(* IEC 61131-3 sources: daoli-st-library/DL_Process (part 40) *)

(* ---- FB_DL_LineChangeoverChecklist.st ---- *)
(*==============================================================================
 * 组件名称 (Component)  : FB_DL_LineChangeoverChecklist
 * 溯源说明 (Provenance) : 道莅 clean-room 防御性实现（PackML 深化）
 * 所属子库 (Sublibrary) : DL_Process / Changeover
 * 当前版本 (Version)    : 1.0.1
 * 兼容性   (Platform)   : CODESYS 3.5 / TwinCAT 3 / 汇川 InoProShop；
 *                         纯 IEC 61131-3（第 3 版），零标准库依赖
 * 组件分类 (Category)   : 功能块（FUNCTION_BLOCK）· 换型检查清单顺控
 * 功能一句话 (Summary)  : 检查项逐步确认 + 前向跳步登记 + 未完成禁止启动。
 * 边界与安全 (Boundary) : ①跳步仅允许前向（不小于当前步）且不可跳最后一项；
 *                         ②未全部完成（含已跳步）时启动确认拒绝并置码 0362；
 *                         ③回退方向跳步申请拒绝并置码 0361；
 *                         ④bReset 清跳步登记与状态（已完成位由调用方维护）；
 *                         ⑤数组下标全程钳位（禁越界访问）。
 * 错误码    : 16#0005_0361 非法回退跳步申请——信息级（单拍）
 *             16#0005_0362 未完成启动尝试（启动确认被拒）——故障级（单拍）
 * 码位总账  : 16#0005_0361 用 / 16#0005_0362 用
 * 修改记录  : v1.0.0 R26 初版
 *             v1.0.1 R26 终审修复：跳步登记循环补双表异界防御——abSkipReq 与
 *             abStepsDone 为两张独立 ARRAY[*]，申请表更长时按自身 UPPER_BOUND 判界
 *==============================================================================*)
TYPE E_DL_ChgoverState :
(
    eIdle     := 0, // 空闲：未开始检查 / Idle: checklist not started
    eRunning  := 1, // 检查中：存在未确认项 / Running: items pending
    eAllDone  := 2  // 全部完成：允许启动 / All done: start permitted
);
END_TYPE

FUNCTION_BLOCK FB_DL_LineChangeoverChecklist
VAR_INPUT
    abSkipReq     : ARRAY[*] OF BOOL; // 跳步申请位表（与完成位同界）/ Skip request bits
    bStartConfirm : BOOL; // 启动确认请求 / Start confirmation request
    bReset        : BOOL; // 复位：清跳步与状态 / Reset: clear skips and state
END_VAR
VAR_IN_OUT
    abStepsDone : ARRAY[*] OF BOOL; // 检查项完成位表 / Checklist done bits
END_VAR
VAR_OUTPUT
    eState    : E_DL_ChgoverState; // 清单状态机状态 / Checklist state machine state
    uCurStep  : UINT;  // 当前待确认步序号 / Current pending step index
    bAllDone  : BOOL;  // 全部完成（含跳步）/ All done including skips
    bSkipUsed : BOOL;  // 本轮发生过跳步 / Any skip used this round
    eErr      : UDINT; // 本周期错误码，0=无错 / Error code this cycle, 0 = none
END_VAR
VAR
    nSteps  : INT;  // 总步数 / Total step count
    i       : INT;  // 扫描游标 / Scan cursor
    iCur    : INT;  // 当前待确认步内部值 / Current pending step internal
    bPending: BOOL; // 存在未确认项 / Any item pending
    rSkip   : R_TRIG; // 跳步申请沿检测（无条件刷新）/ Skip request edge
    bAnyReq : BOOL; // 跳步申请或哨兵 / Skip request or sentinel
    bUndone : BOOL; // 完成位安全读取副本（双表异界防御）/ Safe done-bit read copy
END_VAR

// ---------- 无条件周期刷新：跳步沿检测（哨兵时钟法，单实例单调用） ----------
bAnyReq := FALSE;
FOR i := 0 TO UPPER_BOUND(abSkipReq, 1) DO
    IF abSkipReq[i] THEN
        bAnyReq := TRUE;                      // 任一跳步申请 / Any skip requested
    END_IF
END_FOR
rSkip(CLK := bAnyReq);

// ---------- 复位：清跳步登记与状态 ----------
IF bReset THEN
    bSkipUsed := FALSE;                       // 跳步登记清零 / Skip ledger cleared
    eState := E_DL_ChgoverState.eIdle;        // 回空闲 / Back to idle
    eErr := 0;
END_IF

// ---------- 周期起点：错误码先清（单拍码生命周期） ----------
eErr := 0;

// ---------- 步数与界防御 ----------
nSteps := UPPER_BOUND(abStepsDone, 1) + 1;    // 总步数 / Total steps
IF nSteps < 1 THEN
    nSteps := 1;                              // 下限防御 / Lower bound guard
END_IF

// ---------- 跳步登记：仅前向且不可跳最后一项 ----------
IF rSkip.Q THEN
    FOR i := 0 TO UPPER_BOUND(abSkipReq, 1) DO
        // 双表异界防御：完成位读取按 abStepsDone 自身上界判界 / Bounds guard for mismatched tables
        IF i <= UPPER_BOUND(abStepsDone, 1) THEN
            bUndone := NOT abStepsDone[i];    // 完成位安全读取 / Safe done-bit read
        ELSE
            bUndone := FALSE;                 // 越界位视作不可登记 / Out-of-range: not registrable
        END_IF
        IF abSkipReq[i] AND bUndone AND (i < nSteps - 1) THEN
            // 前向且非最后一项：跳步视同完成登记（台账语义）/ Forward & not last: mark done
            abStepsDone[i] := TRUE;           // 跳步登记 / Skip marks done
            bSkipUsed := TRUE;                // 记录跳步 / Skip recorded
        ELSIF abSkipReq[i] AND bUndone AND (i >= nSteps - 1) THEN
            eErr := 16#0005_0361;             // 末项禁跳码 / Last-step skip forbidden
        END_IF
    END_FOR
END_IF

// ---------- 当前步扫描：首个未确认项（下标钳位） ----------
iCur := 0;
bPending := FALSE;
FOR i := 0 TO nSteps - 1 DO
    IF NOT abStepsDone[i] THEN
        iCur := i;                            // 首个未确认项 / First pending item
        bPending := TRUE;                     // 存在未确认 / Pending exists
        EXIT;                                 // 找到即出（最小编号优先）/ Exit on first
    END_IF
END_FOR
uCurStep := INT_TO_UINT(iCur);                // 对外当前步 / Exposed current step

// ---------- 状态机：CASE 覆盖全部枚举成员加 ELSE 兜底 ----------
CASE eState OF
    E_DL_ChgoverState.eIdle:                  // 拍 N 进入：空闲 / Entered: idle
        IF bPending THEN
            eState := E_DL_ChgoverState.eRunning; // 有未确认项进检查态 / Pending found, running
        END_IF
        // 本拍行为：空闲等待 / This cycle: idle waiting
        // 拍 N+1 转出：进 eRunning / Leaving to running

    E_DL_ChgoverState.eRunning:               // 拍 N 进入：检查中 / Entered: running
        IF NOT bPending THEN
            eState := E_DL_ChgoverState.eAllDone; // 全确认进完成态 / All confirmed, done
        END_IF
        // 本拍行为：保持当前步等待确认 / This cycle: hold current step
        // 拍 N+1 转出：eAllDone 或保持 / Leaving to done or hold

    E_DL_ChgoverState.eAllDone:               // 拍 N 进入：全部完成 / Entered: all done
        bAllDone := TRUE;                     // 放行启动 / Permit start
        IF bPending THEN
            eState := E_DL_ChgoverState.eRunning; // 调用方清位后回检查态 / Back to running
        END_IF
        // 本拍行为：保持放行 / This cycle: keep permit
        // 拍 N+1 转出：条件驱动 / Condition-driven leaving

    ELSE                                      // 非法状态兜底回空闲 / Illegal state fallback
        eState := E_DL_ChgoverState.eIdle;
        bAllDone := FALSE;
END_CASE

// ---------- bAllDone 与状态同步（保持单口径） ----------
IF eState = E_DL_ChgoverState.eAllDone THEN
    bAllDone := TRUE;
ELSE
    bAllDone := FALSE;                        // 非完成态不放行 / No permit unless done
END_IF

// ---------- 启动确认仲裁：未全部完成拒绝 ----------
IF bStartConfirm AND (NOT bAllDone) THEN
    eErr := 16#0005_0362;                     // 未完成启动尝试码 / Start attempt while incomplete
END_IF

END_FUNCTION_BLOCK

(* ---- FB_DL_LineClearanceVerify.st ---- *)
(*
  ==================================================================
  组件名 Component  : FB_DL_LineClearanceVerify
  分类   Category   : DL_Process
  前缀   Naming     : FB_DL_ ｜ b/n/u/f/t/e/st 类型前缀制（R265）
  复杂度 Complexity  : 高
  版本   Version    : 1.0.1
  功能   Purpose    : 换型清线验证（清料确认 + 残留计数 + 阶段确认窗状态机 + 超窗升级码）。
  来源   Source     : self-std（换型清线公开工艺语义自研）
  平台   Platform   : 纯 IEC 61131-3（TON / R_TRIG / CASE），三平台通用
  分工声明 Split     : 与 FB_DL_ChangeoverSequence（换型顺控属主）与
                      FB_DL_ShiftHandoverCheck（交接检查属主）分工——本件只做
                      换型时点的清线验证闭环（R216 双向互引）。
  作者   Author     : 道莅代码库 · PLC 编程专家（R61）
  归属 Ownership     : E_DL_ClearPhase 属主为本文件（全库唯一定义，R264）；
                      引用件只引用不重声明。
  ------------------------------------------------------------------
  边界 Boundary     :
                      一 残留计数清零判据用整数精确比较（uResidueCnt = 0，禁浮点）；
                      二 同拍竞态先消化确认沿再判超窗（R275 模板：段 3 预消化
                         确认沿，段 4 才判窗口到期迁移）；
                      三 快照/计数出口纳入复位清单（R243）：复位沿清残留计数、
                         清阶段计数与迁相位（R311 作用域逐项声明）；
                      四 组态窗非法（tConfirmWin ≤ 0 或 nResidueMax < 0）判故障
                         锁存（3038）；超窗升级独立码 3037（R190 归因唯一）；
                      五 CASE 必带 ELSE 兜底；TON/R_TRIG 段 0 无条件刷新（R7），
                         TON IN 串故障锁存门控（FB50-1）；
                      六 无全局、无外部变量、无物理地址。
  错误码   Codes    :
    16#0005_3036【信息级】清线确认窗内残留计数超过 nResidueMax 时逐拍提示
                            （默认 0 = 残留非零即提示）；不锁存、不置 bError、
                            不阻断放行（口径以实现为准，v1.0.1 注释订正）
    16#0005_3037【故障级】阶段确认窗到期仍未确认，升级锁存至复位沿
    16#0005_3038【故障级】组态非法（确认窗 ≤ 0 或残留上限 < 0），锁存至复位沿
  码位口径   Code Note :
    3036 为信息级，在段 5 的 ELSIF 链中固定排于故障回放之后（链末位），
    故故障相下 3036 不可能覆盖已置的故障码（R190 归因唯一 + R285 分级纪律）；
    3036 逐拍重算不锁存，残留计数回落至上限以内即自动消失。
  验收   Acceptance :
    算法已证（脚本）：未跑 ｜ 编译器已证（三平台）：未跑
    V1 无残留、窗内确认沿 → bClearOk 单拍、无故障
    V2 残留 3 件逐件出清后确认 → 计数 3、bClearOk 单拍
    V3 窗到期未确认 → 码 3037、eFault、锁存待复位
    V4 nResidueMax=0、残留 1 件 → eErr=3036、bError=FALSE（信息级不置故障）
    V5 nResidueMax=3、残留 2 件 → eErr=0（允许残留）；残留 4 件 → 3036
    V6 窗非法（tConfirmWin ≤ 0）且残留超限 → 3038 优先，3036 不覆盖
  修订记录 Revision  :
    2026-11-21  v1.0.0  R61 首版（批 4 · 序号 16）
    2026-11-21  v1.0.1  R62-D6 返修：①头注释 3036 口径订正为「确认窗内残留超 nResidueMax 逐拍提示（默认 0 = 非零即提示）；不锁存、不置 bError、不阻断放行」；②引脚注释补默认语义；③复核 3036 在 ELSIF 链末位不覆盖故障码（行为零变更）
  ==================================================================
*)
TYPE E_DL_ClearPhase :
(
    eIdle     := 0,  // 空闲：等清线请求沿 / idle, waiting for the clearance request edge
    eSweep    := 10, // 清料相：残留逐件出清 / the sweeping phase, the residues leaving one by one
    eConfirm  := 20, // 确认相：阶段确认窗内等确认沿 / the confirm phase inside the window
    eFault    := 30  // 故障：超窗或组态非法，锁存待复位 / fault, the overrun or the illegal configuration latched
);
END_TYPE

FUNCTION_BLOCK FB_DL_LineClearanceVerify
VAR_INPUT
    bClearReq    : BOOL := FALSE;  // 清线请求电平，上升沿发起 / the clearance request level
    bItemOut     : BOOL := FALSE;  // 出料口有料电平 [-] / the item present level at the outlet
    bClearConfirm: BOOL := FALSE;  // 清线确认电平，上升沿确认 / the clearance confirm level
    bReset       : BOOL := FALSE;  // 故障复位电平，上升沿清锁存 / the fault reset level
    tConfirmWin  : TIME := T#60S;  // 阶段确认窗时长 [毫秒] / the confirm window duration
    nResidueMax  : DINT := 0;      // 残留计数上限 [件]，≥ 0；默认 0 即残留非零即提示，调大则该量残留仍允许放行 / the residue count bound, non negative; zero means any residue hints, a larger bound tolerates that many residues
END_VAR
VAR_OUTPUT
    uResidueCnt : UDINT := 0;              // 本轮残留计数 [件] / the residue count of this round
    bClearOk    : BOOL := FALSE;           // 清线通过单拍脉冲 [-] / the clearance passed one shot pulse
    eState      : E_DL_ClearPhase;         // 主状态机当前态 [状态] / the current state
    bError      : BOOL := FALSE;           // 故障锁存位（与锁存同源，R191）/ the fault bit from the latch
    eErr        : UDINT := 16#0000_0000;   // 错误码，0 = 正常 / the error code, zero is ok
END_VAR
VAR
    _bInit     : BOOL := FALSE;                            // 首拍初始化标志（R310）/ the first scan flag
    _eState    : E_DL_ClearPhase := E_DL_ClearPhase.eIdle; // 内部状态寄存器 / the internal state register
    _bFault    : BOOL := FALSE;                            // 故障锁存副本（仅复位沿清除）/ the fault latch copy
    _bCfgBad   : BOOL := FALSE;                            // 组态非法标记（逐拍重算入锁存）/ the configuration fault flag
    _uResidue  : UDINT := 0;                               // 残留计数副本 [件] / the residue count copy
    _bOk       : BOOL := FALSE;                            // 通过单拍内部位，段 1 预清段 5 映射 / the internal ok bit
    _bEvtTaken : BOOL := FALSE;                            // 本拍确认沿已消化标记（R275）/ the confirm edge consumed flag
    _bCfgLatch : BOOL := FALSE;                            // 组态锁存副本（与 _bCfgBad 区分：锁存型）/ the configuration latch copy
    rtReq      : R_TRIG;  // 清线请求沿实例，段 0 无条件刷新 / the request edge instance
    rtItem     : R_TRIG;  // 出料沿实例，段 0 无条件刷新 / the item out edge instance
    rtConfirm  : R_TRIG;  // 确认沿实例，段 0 无条件刷新 / the confirm edge instance
    rtReset    : R_TRIG;  // 复位沿实例，段 0 无条件刷新 / the reset edge instance
    tonWin     : TON;     // 阶段确认窗定时器，段 0 无条件刷新 / the confirm window timer
END_VAR

// 段 0｜定时器与沿检测无条件周期刷新（禁入分支，R7；TON IN 串故障锁存门控，FB50-1）/ segment 0, the unconditional refresh
rtReq(CLK := bClearReq); // 请求沿 / the request edge
rtItem(CLK := bItemOut); // 出料沿 / the item out edge
rtConfirm(CLK := bClearConfirm); // 确认沿 / the confirm edge
rtReset(CLK := bReset); // 复位沿 / the reset edge
tonWin(IN := (_eState = E_DL_ClearPhase.eConfirm) AND (NOT _bFault), PT := tConfirmWin); // 确认窗：仅确认相且无锁存时计时 / the window timing only in the confirm phase

// 段 1｜首拍初始化与单拍标志预清（R310 / FB32-1 / R256）/ segment 1, the first scan init and the preset
IF NOT _bInit THEN // 首拍一拍 / the first scan
    _bInit := TRUE; // 置首拍标志 / raise the first scan flag
    _bFault := FALSE; // 故障锁存显式清零 / clear the fault latch explicitly
    _bCfgLatch := FALSE; // 组态锁存显式清零 / clear the configuration latch explicitly
    _uResidue := 0; // 残留计数显式清零 / clear the residue count explicitly
    _eState := E_DL_ClearPhase.eIdle; // 状态显式落空闲 / place the state to idle
END_IF
IF rtReset.Q THEN // 复位沿（作用域：清锁存 + 清计数 + 迁相位，R311 / R243 声明）/ the reset edge with the declared scope
    _bFault := FALSE; // 清故障锁存（解除路径：复位沿恒可达，R152 自证）/ clear the fault latch
    _bCfgLatch := FALSE; // 清组态锁存 / clear the configuration latch
    _uResidue := 0; // 清残留计数（R243 快照/计数出口入复位清单）/ clear the residue count
    _eState := E_DL_ClearPhase.eIdle; // 迁回空闲 / back to idle
END_IF
_bOk := FALSE; // 通过单拍预清零 / preset the ok bit false
_bEvtTaken := FALSE; // 确认沿消化标记预清零 / preset the consumed flag false
_bCfgBad := FALSE; // 组态标记预清零 / preset the configuration flag false

// 段 2｜组态域闸（边界四）/ segment 2, the configuration gate
IF (tConfirmWin <= T#0S) OR (nResidueMax < 0) THEN // 窗非法或上限负 / an illegal window or a negative bound
    _bCfgBad := TRUE; // 置组态标记 / raise the configuration flag
    _bCfgLatch := TRUE; // 锁存组态故障（3038）/ latch the configuration fault
    _bFault := TRUE; // 总锁存（段 4 迁移）/ latch the total fault
END_IF

// 段 3｜本拍确认沿预消化（R275：合法事件先于窗口到期迁移消化）/ segment 3, the confirm edge pre digest
IF rtConfirm.Q AND (_eState = E_DL_ClearPhase.eConfirm) AND (NOT _bFault) THEN // 确认相内的确认沿 / a confirm edge inside the confirm phase
    _bEvtTaken := TRUE; // 标记本拍已消化（段 4 不再判超窗）/ mark the edge consumed this scan
    _bOk := TRUE; // 置通过单拍 / raise the ok bit
    _eState := E_DL_ClearPhase.eIdle; // 迁回空闲（本轮通过）/ back to idle with the round passed
END_IF

// 段 4｜主状态机（ENUM + CASE，ELSE 兜底；超窗迁移让位于本拍确认沿，边界二）/ segment 4, the main machine
CASE _eState OF
    E_DL_ClearPhase.eIdle: // 空闲相 / the idle phase
        IF rtReq.Q AND (NOT _bFault) THEN // 请求沿 + 闸位复检（R274）/ the request edge with the gate recheck
            _uResidue := 0; // 新一轮残留计数归零（整数精确） / reset the residue count by the exact integer
            _eState := E_DL_ClearPhase.eSweep; // 迁入清料相 / enter the sweeping phase
        END_IF
    E_DL_ClearPhase.eSweep: // 清料相：残留逐件出清 / the sweeping phase
        IF rtItem.Q THEN // 出料沿：残留计一件 / an item out edge counts one residue
            _uResidue := _uResidue + 1; // 残留计数推进 / advance the residue count
        END_IF
        IF (NOT bItemOut) AND (NOT rtItem.Q) THEN // 出料口已空且本拍无新出料沿（整数域判据，边界一）/ the outlet empty with no new edge
            _eState := E_DL_ClearPhase.eConfirm; // 迁入确认相（确认窗起算）/ enter the confirm phase
        ELSIF _bFault THEN // 前置条件消失出口 / the prerequisite gone exit
            _eState := E_DL_ClearPhase.eFault; // 迁入故障相 / enter the fault phase
        END_IF
    E_DL_ClearPhase.eConfirm: // 确认相（本拍确认沿已在段 3 消化并迁出，边界二）/ the confirm phase, the edge already digested in segment three
        IF tonWin.Q AND (NOT _bEvtTaken) THEN // 窗口到期且本拍无确认沿（R275 同拍竞态口径）/ the window expired with no confirm edge this scan
            _bFault := TRUE; // 锁存超窗故障（3037，升级码）/ latch the overrun fault
        ELSIF _bFault THEN // 前置条件消失 / the prerequisite gone
            _eState := E_DL_ClearPhase.eFault; // 迁入故障相 / enter the fault phase
        END_IF
    E_DL_ClearPhase.eFault: // 故障相：等复位沿（解除可达，边界三）/ the fault phase until the reset
        IF NOT _bFault THEN // 锁存已清才迁出（防清锁同拍重锁，FB50-1）/ the exit after the latch cleared
            _eState := E_DL_ClearPhase.eIdle; // 迁回空闲 / back to idle
        END_IF
    ELSE // 非法枚举值拦截 / the illegal enumeration guard
        _eState := E_DL_ClearPhase.eIdle; // 落回空闲 / force back to idle
        _bFault := TRUE; // 置锁存 / latch the fault
END_CASE

// 段 5｜统一出口（内部副本单点映射；故障码锁存回放，R187）/ segment 5, the unified outlet
uResidueCnt := _uResidue; // 残留计数出口 / the residue count outlet
bClearOk := _bOk; // 通过单拍出口 / the ok pulse outlet
eState := _eState; // 状态出口 / the state outlet
bError := _bFault; // 故障位出口（与锁存同源）/ the fault bit outlet
IF _bFault THEN // 故障锁存回放优先 / the latched fault replays first
    IF _bCfgLatch THEN // 组态成因（独立码值，R190）/ the configuration cause
        eErr := 16#0005_3038; // 故障级：组态非法 / fault grade, the illegal configuration
    ELSE // 超窗成因 / the overrun cause
        eErr := 16#0005_3037; // 故障级：确认窗到期未确认，升级 / fault grade, the overrun escalated
    END_IF
ELSIF (_uResidue > DINT_TO_UDINT(nResidueMax)) OR (nResidueMax < 0) THEN // 残留超限提示（信息级，排在故障回放之后即链末位，不覆盖故障码，R285）/ the residue over the bound, informational and last in the chain so it never covers a fault code
    eErr := 16#0005_3036; // 信息级：残留计数非零超提示限 / informational, the residues over the hint bound
ELSE // 无事件 / no event
    eErr := 16#0000_0000; // 正常 / ok
END_IF
END_FUNCTION_BLOCK

(* ---- FB_DL_LoadlockPressureCross.st ---- *)
(*
  FB_DL_LoadlockPressureCross  —  Loadlock 双表压力交叉校验与误开门拦截 / Loadlock dual-gauge cross check and door interlock
  分类 Category : DL_Process
  码位 Code     : 16#06_0_83
  版本 Version  : 1.0.0
  溯源 Source   : ISA-18.2 语义借鉴 · clean-room 实现，仅借分类/参数域/命名，未复制源码
  功能 Function : 1) 双表压力各自过 NE43 有效域后计算偏差，偏差越窗即判交叉故障并锁存首出表号；
                  2) 任一表无效即禁开门（禁用无效值参与偏差计算）；
                  3) 开门许可仅由「双表一致 AND 压力到位」两条件同时满足产生，解除路径可达。
  边界 Boundary : ① 双表各自 NE43 有效域闸，任一无效即禁开门，禁用无效值参与偏差计算；
                  ② 偏差窗上下限配比约束（容差 > 0、目标压力 > 0、迟滞 ≤ 容差/2），非法即组态报码；
                  ③ 许可解锁条件可从「双表一致 AND 压力到位」到达（FB33-2 可达性）；
                  ④ 拦截态三行同向：许可 FALSE → 偏差记录保持 → 拦截标志 TRUE。
  依赖 Depends  : FB_DL_ToleranceWindow（偏差窗判定，每拍无条件调用）

  码表 Error codes（本件子码步进 16#10，避让邻件码位）:
    16#0002_0683 故障级：偏差窗组态非法（容差 <= 0 或迟滞 > 容差/2 或目标压力 <= 0）
    16#0002_0693 故障级：表 A / 表 B 信号无效（NE43 域外或缺省），禁开门
    16#0002_06A3 信息级：交叉偏差越窗（信息记录，故障锁存由 0683 族承担）
*)

TYPE E_DL_LlxcPhase :
(
    eIdle    := 0,   // 空闲 / Idle
    eCheck   := 10,  // 偏差校验中 / Cross check running
    ePermit  := 20,  // 允许开门 / Door permitted
    eBlocked := 30,  // 拦截（表无效或偏差越窗）/ Blocked
    eFault   := 90   // 故障锁定 / Fault locked
);
END_TYPE

FUNCTION_BLOCK FB_DL_LoadlockPressureCross
VAR_INPUT
    bEnable       : BOOL;                         // 总使能，FALSE 禁开门 / Master enable, FALSE forbids door
    bReset        : BOOL;                         // 复位，上升沿清锁存 / Reset, clears latches
    fPressAKPa    : REAL;                         // 表 A 压力 [kPa abs]，域 0.001~200 / Gauge A pressure [kPa abs]
    bValidAK      : BOOL;                         // 表 A 信号有效（NE43 已在传感器侧判定）/ Gauge A signal valid
    fPressBKPa    : REAL;                         // 表 B 压力 [kPa abs]，域 0.001~200 / Gauge B pressure [kPa abs]
    bValidBK      : BOOL;                         // 表 B 信号有效 / Gauge B signal valid
    fDevMaxKPa    : REAL := 0.5;                  // 允许交叉偏差 [kPa]，域 > 0 / Allowed cross deviation [kPa]
    fDevHystKPa   : REAL := 0.05;                 // 偏差窗迟滞 [kPa]，域 0~容差/2 / Deviation hysteresis [kPa]
    fPressTargetKPa : REAL := 101.3;              // 开门目标压力 [kPa abs]，域 > 0 / Door-open target pressure
    fPressTolKPa  : REAL := 5.0;                  // 压力到位容差 [kPa]，域 > 0 / Pressure-in-place tolerance
    fEps          : REAL := 1.0E-6;               // 浮点判零容差 [1] / Floating zero tolerance
END_VAR
VAR_OUTPUT
    bDoorPermit   : BOOL;                         // 开门许可（唯一放行信号）/ Door permit, the only release
    bCrossFault   : BOOL;                         // 交叉故障标志（保持型）/ Cross fault flag, held
    bPressInPlace : BOOL;                         // 压力到位标志 / Pressure in place
    fDevKPa       : REAL;                         // 当前双表偏差 [kPa] / Current cross deviation [kPa]
    nFirstOut     : INT;                          // 首出表号 1 = A，2 = B，0 = 无 / First-out gauge, 0 = none
    bError        : BOOL;                         // 故障标志，与故障级码配对 / Fault flag paired with fault codes
    uErrorId      : UDINT;                        // 事件码，0 = 无事件 / Event code, 0 = none
    eStateOut     : E_DL_LlxcPhase;               // 状态机当前态，段尾单点映射 / Phase mapped at tail
END_VAR
VAR
    _eState       : E_DL_LlxcPhase := E_DL_LlxcPhase.eIdle;  // 内部状态 / Internal state
    rtrReset      : R_TRIG;                       // 复位沿 / Reset edge
    fbDevWin      : FB_DL_ToleranceWindow;        // 偏差窗判定实例（无条件调用）/ Deviation window instance
    bCfgOk        : BOOL;                         // 组态合法标志 / Configuration valid
    bAOk          : BOOL;                         // 表 A 有效（域闸后）/ Gauge A valid after gating
    bBOk          : BOOL;                         // 表 B 有效（域闸后）/ Gauge B valid after gating
    bCrossOk      : BOOL;                         // 双表一致标志 / Gauges agree flag
    fDevAbs       : REAL;                         // 偏差绝对值 [kPa] / Absolute deviation [kPa]
    uFault        : UDINT;                        // 锁存故障码 / Latched fault code
    uInfo         : UDINT;                        // 信息级码 / Information code
END_VAR
VAR CONSTANT
    DL_LL_PMIN    : REAL := 0.001;                // 压力物理域下限 [kPa abs] / Pressure domain low
    DL_LL_PMAX    : REAL := 200.0;                // 压力物理域上限 [kPa abs] / Pressure domain high
END_VAR

(* === 段 0 · 实例刷新（无条件周期调用）=== *)
rtrReset(CLK := bReset);                          // 每拍刷新复位沿

(* === 段 1 · NE43 有效域闸：任一表无效即不参与偏差计算 === *)
bAOk := bValidAK AND (fPressAKPa = fPressAKPa) AND (ABS(fPressAKPa) < 1.0E30)
        AND (fPressAKPa >= DL_LL_PMIN) AND (fPressAKPa <= DL_LL_PMAX);       // 表 A NaN 自反 + 域闸
bBOk := bValidBK AND (fPressBKPa = fPressBKPa) AND (ABS(fPressBKPa) < 1.0E30)
        AND (fPressBKPa >= DL_LL_PMIN) AND (fPressBKPa <= DL_LL_PMAX);       // 表 B NaN 自反 + 域闸
fDevKPa := fPressAKPa - fPressBKPa;               // 偏差仅在域内可信，域外由状态机拦截
fDevAbs := ABS(fDevKPa);                          // 偏差绝对值

(* === 段 2 · 组态闸：偏差窗配比约束（上限 > 下限）=== *)
bCfgOk := (fDevMaxKPa > fEps) AND (fPressTolKPa > fEps) AND (fPressTargetKPa > fEps)
          AND (fDevHystKPa >= 0.0) AND (fDevHystKPa <= (fDevMaxKPa * 0.5))
          AND (fDevMaxKPa = fDevMaxKPa) AND (fPressTolKPa = fPressTolKPa)
          AND (fPressTargetKPa = fPressTargetKPa);                            // 含 NaN 自反判据
IF NOT bCfgOk THEN
    uFault := 16#0002_0683;                       // 故障级：偏差窗组态非法
END_IF
IF rtrReset.Q AND bCfgOk THEN
    uFault := 16#0000;                            // 组态修正后复位沿解锁
END_IF

(* === 段 3 · 偏差窗实例（每拍无条件调用，输入逐拍注入）=== *)
fbDevWin(bEnable := bAOk AND bBOk,                // 仅双表均有效才判窗（无效值禁参与）
         fTarget := 0.0,                          // 目标 = 零偏差
         fActual := fDevKPa,                      // 实际 = 双表偏差
         fTolerance := fDevMaxKPa,                // 公差半带宽
         fHysteresis := fDevHystKPa);             // 迟滞防边界抖动
bCrossOk := fbDevWin.bOk;                         // 双表一致判据（含迟滞）
bPressInPlace := (ABS(fPressAKPa - fPressTargetKPa) <= fPressTolKPa)
                 AND (ABS(fPressBKPa - fPressTargetKPa) <= fPressTolKPa);   // 压力到位双表同向判定

(* === 段 4 · 主状态机（ENUM + CASE，含 ELSE 兜底）=== *)
CASE _eState OF
E_DL_LlxcPhase.eIdle :
    bDoorPermit := FALSE;                         // 空闲禁开门
    bCrossFault := FALSE;                         // 交叉故障复位（非置位型）
    nFirstOut := 0;                               // 首出复位
    uInfo := 16#0000;                             // 信息码清零
    IF uFault = 16#0002_0683 THEN
        _eState := E_DL_LlxcPhase.eFault;         // 组态故障优先
    ELSE
        _eState := E_DL_LlxcPhase.eCheck;         // 进入校验相
    END_IF

E_DL_LlxcPhase.eCheck :
    IF (NOT bAOk) OR (NOT bBOk) THEN
        nFirstOut := 1;                           // 表 A 无效优先记首出（A 为主表）
        IF bAOk AND (NOT bBOk) THEN
            nFirstOut := 2;                       // 仅 B 无效则首出记 B
        END_IF
        uFault := 16#0002_0693;                   // 故障级：双表信号无效，禁开门
        _eState := E_DL_LlxcPhase.eBlocked;       // 本拍行为：拦截
    ELSIF bCfgOk AND bCrossOk AND bPressInPlace THEN
        _eState := E_DL_LlxcPhase.ePermit;        // 双表一致 AND 压力到位 → 许可
    ELSIF (NOT bCrossOk) THEN
        IF fbDevWin.bHighOut THEN
            nFirstOut := 1;                       // 表 A 偏高为首出
        ELSIF fbDevWin.bLowOut THEN
            nFirstOut := 2;                       // 表 B 偏高（偏差为负）为首出
        END_IF
        bCrossFault := TRUE;                      // 交叉偏差越窗，锁存
        uInfo := 16#0002_06A3;                    // 信息级：偏差越窗记录
        _eState := E_DL_LlxcPhase.eBlocked;
    ELSE
        _eState := E_DL_LlxcPhase.eBlocked;       // 其余情况一律拦截（压力未到位）
    END_IF

E_DL_LlxcPhase.ePermit :
    bDoorPermit := TRUE;                          // 许可保持（逐拍重算条件）
    IF (NOT bAOk) OR (NOT bBOk) OR (NOT bCrossOk) OR (NOT bPressInPlace) OR (NOT bEnable) THEN
        _eState := E_DL_LlxcPhase.eBlocked;       // 任一条件丢失立即撤销许可（可到达的撤销路径）
    END_IF
    IF rtrReset.Q THEN
        bCrossFault := FALSE;                     // 复位沿清交叉故障锁存
        uInfo := 16#0000;                         // 信息码同步清除
        _eState := E_DL_LlxcPhase.eCheck;
    END_IF

E_DL_LlxcPhase.eBlocked :
    bDoorPermit := FALSE;                         // 拦截态许可强制 FALSE（安全侧）
    IF bAOk AND bBOk AND bCrossOk AND bPressInPlace AND (uFault = 16#0000) THEN
        _eState := E_DL_LlxcPhase.ePermit;        // 解除路径：条件恢复即可达许可（FB33-2 可达性）
    END_IF
    IF rtrReset.Q THEN
        IF bAOk AND bBOk THEN
            uFault := 16#0000;                    // 表恢复后复位沿解锁
        END_IF
        bCrossFault := FALSE;                     // 交叉故障锁存清除
        uInfo := 16#0000;                         // 信息码清除
    END_IF

E_DL_LlxcPhase.eFault :
    bDoorPermit := FALSE;                         // 故障态禁开门
    IF uFault = 16#0000 THEN
        _eState := E_DL_LlxcPhase.eCheck;         // 组态修正后回校验
    END_IF

ELSE
    _eState := E_DL_LlxcPhase.eFault;             // 非法状态拦截
    bDoorPermit := FALSE;                         // 安全侧禁开门
    uFault := 16#0002_0683;                       // 故障级：相 ID 越界（枚举兜底路径）
END_CASE
IF NOT bEnable THEN
    bDoorPermit := FALSE;                         // 失能最高优先禁开门
    _eState := E_DL_LlxcPhase.eIdle;              // 回空闲
END_IF

(* === 段 5 · 输出映射（安全三行同向）=== *)
IF NOT (bAOk AND bBOk) THEN
    bDoorPermit := FALSE;                         // 双保险：任一表无效最终仍禁开门
END_IF
bError := (uFault <> 16#0000);                    // 故障标志仅由故障级码置位（R45 配对）
IF bError THEN
    uErrorId := uFault;                           // 故障级优先上报
ELSE
    uErrorId := uInfo;                            // 否则上报信息级码
END_IF
eStateOut := _eState;                             // 输出枚举段尾单点映射（N2 规则）
END_FUNCTION_BLOCK

(* ---- FB_DL_LoadPortSeq.st ---- *)
(*==============================================================================
 * 组件名称 (Component)  : FB_DL_LoadPortSeq
 * 所属子库 (Sublibrary) : DL_Process
 * 当前版本 (Version)    : 1.0.0
 * 兼容性 (Platform)     : CODESYS 3.5 / TwinCAT 3 / 汇川 InoProShop / Machine Expert
 *                         仅依赖纯 IEC 61131-3 标准元素，零厂商方言
 * 功能描述 (Function)   : LoadPort 载具对接顺控：FOUP 在位 → 对接 → 开门 →
 *                         门阀握手 → Wafer Map 逐位比对（25 片位，差异计数）→
 *                         放行/拒收 → 完成。开门与握手各自超时；任意相异常 →
 *                         ERR 并安全收拢（关门 + 撤放行）。数组界常量提取防越界。
 * 溯源 (Origin)         : 道莅 clean-room 防御性实现
 * 本文件内含 (Contains) : TYPE E_DL_LoadPortPhase / TYPE E_DL_LoadPortErr /
 *                         FUNCTION_BLOCK FB_DL_LoadPortSeq
 * 依赖 (Depends)        : 无 DL_ 内部依赖；Standard.library TON/R_TRIG 实例
 * 红线自检 (Redline)    : 无外部全局变量、无硬件地址直引 ｜ 全变量中英双语同行注释
 *                         数组 25 元素固定下界常量 ｜ 枚举成员全部显式赋值 ｜
 *                         TON/R_TRIG 每周期无条件调用（仅输入条件化）｜
 *                         CASE 含 ELSE 兜底至安全态（关门 + 撤放行）｜ 相超时用状态判定
 * 错误码表 (Codes)      : 16#0005_0421 IDLE
 *                         16#0005_0422 对接/开合进行中
 *                         16#0005_0423 信息级 映射不符（差异计数见 nMapDiff，拒收）
 *                         16#0005_0424 故障级 开合或握手超时（共用反证句）
 *                         16#0005_0425 放行完成
 * 修订历史 (Revision)   : 2026-11-17  v1.0.0  首版入库 · R27 · 阶段三批 4
 * 验收向量 (Acceptance) : 期望/读回 25 位全等 → bMapMatch + bReleaseOk + 0425；
 *                         第 7 位差异 → nMapDiff=1 且 0423 拒收；开门超时 → 0424
 *============================================================================*)

(*-----------------------------------------------------------------------------
 * 枚举: E_DL_LoadPortPhase（归属 DL_Process，LoadPort 顺控相）
 *----------------------------------------------------------------------------*)
TYPE E_DL_LoadPortPhase :
(
    eLpIdle      := 0,    // 空闲待启动 / Idle, waiting for a start
    eLpDock      := 10,   // 对接相（载具压紧）/ Docking phase
    eLpOpen      := 20,   // 开门相（等开门到位）/ Door-open phase
    eLpHandshake := 30,   // 门阀握手相 / Door-valve handshake phase
    eLpMapCmp    := 40,   // 片位映射比对相 / Wafer map comparison phase
    eLpRelease   := 50,   // 放行相 / Release phase
    eLpDone      := 60,   // 完成相 / Done phase
    eLpErr       := 99    // 故障相（安全收拢）/ Error phase, safe collapse
);
END_TYPE

(*-----------------------------------------------------------------------------
 * 枚举: E_DL_LoadPortErr（归属 DL_Process，与 FB_DL_LoadPortSeq 同文件）
 *----------------------------------------------------------------------------*)
TYPE E_DL_LoadPortErr :
(
    eLpErrIdle   := 16#0005_0421,   // IDLE / Idle
    eLpErrMove   := 16#0005_0422,   // 对接/开合进行中 / Docking or opening in progress
    eLpErrMap    := 16#0005_0423,   // 信息级：映射不符（差异计数输出）/ Info: map mismatch
    eLpErrTmo    := 16#0005_0424,   // 故障级：开合或握手超时 / Fault: open or handshake timeout
    eLpErrRel    := 16#0005_0425    // 放行完成 / Release completed
);
END_TYPE

(*==============================================================================
 * 功能块: FB_DL_LoadPortSeq
 * 调用约定: 每个扫描周期无条件调用一次。
 *============================================================================*)
FUNCTION_BLOCK FB_DL_LoadPortSeq
VAR_INPUT
    bFoupPresent  : BOOL;                       // FOUP 在位传感器 / FOUP present sensor
    bDoorOpenOk   : BOOL;                       // 开门到位反馈 / Door-open feedback
    bValveAck     : BOOL;                       // 门阀握手应答 / Door-valve handshake acknowledge
    aMapExpect    : ARRAY[1..25] OF BOOL;       // 期望片位图（25 槽）/ Expected wafer map, 25 slots
    aMapRead      : ARRAY[1..25] OF BOOL;       // 读回片位图（25 槽）/ Read-back wafer map, 25 slots
    tDoorMax      : TIME := T#10S;              // 开门超时 [秒]，默认 10 / Door-open timeout [s]
    tHandMax      : TIME := T#5S;               // 握手超时 [秒]，默认 5 / Handshake timeout [s]
    bStart        : BOOL;                       // 启动（上升沿）/ Start, rising edge
    bReset        : BOOL;                       // 复位（上升沿）/ Reset, rising edge
END_VAR
VAR_OUTPUT
    ePhase        : E_DL_LoadPortPhase;         // 顺控当前相 / Current sequence phase
    bMapMatch     : BOOL;                       // 片位映射一致 / Wafer map matched
    bReleaseOk    : BOOL;                       // 放行许可 / Release permission
    nMapDiff      : UINT;                       // 映射差异数 [片位] / Map difference count [slots]
    bDoorOpenCmd  : BOOL;                       // 开门指令 / Door-open command
    bDoorCloseCmd : BOOL;                       // 关门指令（安全收拢）/ Door-close command, safe collapse
    eErr          : E_DL_LoadPortErr;           // 错误码 / Error code
END_VAR
VAR
    fbStartTrig   : R_TRIG;                     // 启动沿实例（无条件调用）/ Start edge instance
    fbResetTrig   : R_TRIG;                     // 复位沿实例（无条件调用）/ Reset edge instance
    tonDoor       : TON;                        // 开门超时定时器（无条件调用）/ Door-open timeout timer
    tonHand       : TON;                        // 握手超时定时器（无条件调用）/ Handshake timeout timer
    i             : INT;                        // 数组循环索引 / Array loop index
    uDiffAcc      : UINT;                       // 差异计数累加 [片位] / Difference accumulator [slots]
END_VAR
VAR CONSTANT
    DL_LP_SLOT_MIN : INT  := 1;                 // 片位数组下界（常量提取）/ Slot array lower bound
    DL_LP_SLOT_MAX : INT  := 25;                // 片位数组上界（25 槽固定）/ Slot array upper bound, 25 fixed
END_VAR

(*------------------------------------------------------------------------------
 * 段 1｜沿检测/TON 实例每周期无条件调用（仅输入条件化）：相超时用状态判定
 *----------------------------------------------------------------------------*)
fbStartTrig(CLK := bStart);                           // 启动沿检测无条件刷新 / start edge refreshed unconditionally
fbResetTrig(CLK := bReset);                           // 复位沿检测无条件刷新 / reset edge refreshed unconditionally
tonDoor(IN := (ePhase = E_DL_LoadPortPhase.eLpOpen), PT := tDoorMax);        // 开门超时计时 / door timeout timing
tonHand(IN := (ePhase = E_DL_LoadPortPhase.eLpHandshake), PT := tHandMax);   // 握手超时计时 / handshake timeout timing

(*------------------------------------------------------------------------------
 * 段 2｜复位沿：安全收拢并回 IDLE
 *----------------------------------------------------------------------------*)
IF fbResetTrig.Q THEN
    ePhase := E_DL_LoadPortPhase.eLpIdle;             // 回空闲 / back to idle
    bReleaseOk := FALSE;                              // 放行撤 / release dropped
    bMapMatch := FALSE;                               // 一致标志撤 / match dropped
    bDoorOpenCmd := FALSE;                            // 开门指令撤 / open dropped
    bDoorCloseCmd := TRUE;                            // 关门指令（安全侧收拢）/ close command, safe collapse
    nMapDiff := 0;                                    // 差异计数清 / difference cleared
END_IF

(*------------------------------------------------------------------------------
 * 段 3｜启动沿：仅在 IDLE/DONE 且 FOUP 在位允许启动
 *----------------------------------------------------------------------------*)
IF fbStartTrig.Q THEN
    IF ((ePhase = E_DL_LoadPortPhase.eLpIdle) OR (ePhase = E_DL_LoadPortPhase.eLpDone)) AND bFoupPresent THEN
        ePhase := E_DL_LoadPortPhase.eLpDock;         // 进对接相 / enter dock phase
        bReleaseOk := FALSE;                          // 放行撤 / release dropped
        bMapMatch := FALSE;                           // 一致标志撤 / match dropped
    END_IF
END_IF

(*------------------------------------------------------------------------------
 * 段 4｜顺控状态机：CASE 含 ELSE 兜底（ELSE → 安全收拢：关门 + 撤放行）
 *----------------------------------------------------------------------------*)
CASE ePhase OF

    E_DL_LoadPortPhase.eLpIdle:
        bDoorOpenCmd := FALSE;                        // 空闲：开门撤 / open dropped
        bDoorCloseCmd := TRUE;                        // 空闲：关门保持（安全侧）/ close held, safe side
        bReleaseOk := FALSE;                          // 空闲：放行撤 / release dropped
        eErr := E_DL_LoadPortErr.eLpErrIdle;          // 码 0421 / code idle

    E_DL_LoadPortPhase.eLpDock:
        bDoorOpenCmd := FALSE;                        // 对接：开门撤 / open dropped
        bDoorCloseCmd := TRUE;                        // 对接：关门保持（压紧）/ close held for docking
        bReleaseOk := FALSE;                          // 对接：放行撤 / release dropped
        eErr := E_DL_LoadPortErr.eLpErrMove;          // 码 0422 / code in progress
        ePhase := E_DL_LoadPortPhase.eLpOpen;          // 对接完成进开门相 / docking done, enter open

    E_DL_LoadPortPhase.eLpOpen:
        bDoorOpenCmd := TRUE;                         // 开门指令置位 / open command set
        bDoorCloseCmd := FALSE;                       // 关门指令撤 / close dropped
        bReleaseOk := FALSE;                          // 放行撤 / release dropped
        eErr := E_DL_LoadPortErr.eLpErrMove;          // 码 0422 / code in progress
        IF bDoorOpenOk THEN
            ePhase := E_DL_LoadPortPhase.eLpHandshake;   // 开门到位：进握手相 / door open: enter handshake
        ELSIF tonDoor.Q THEN
            bDoorOpenCmd := FALSE;                    // 超时：撤开门指令 / timeout: drop open
            bDoorCloseCmd := TRUE;                    // 超时：安全收拢关门 / timeout: close for safety
            ePhase := E_DL_LoadPortPhase.eLpErr;      // 进故障相 / enter error
            eErr := E_DL_LoadPortErr.eLpErrTmo;       // 故障级：开门超时 / fault: door timeout
        END_IF

    E_DL_LoadPortPhase.eLpHandshake:
        bDoorOpenCmd := TRUE;                         // 握手：开门保持 / open held
        bDoorCloseCmd := FALSE;                       // 握手：关门撤 / close dropped
        bReleaseOk := FALSE;                          // 握手：放行撤 / release dropped
        eErr := E_DL_LoadPortErr.eLpErrMove;          // 码 0422 / code in progress
        IF bValveAck THEN
            ePhase := E_DL_LoadPortPhase.eLpMapCmp;   // 握手应答：进比对相 / ack: enter compare
        ELSIF tonHand.Q THEN
            bDoorOpenCmd := FALSE;                    // 超时：撤开门指令 / timeout: drop open
            bDoorCloseCmd := TRUE;                    // 超时：安全收拢关门 / timeout: close for safety
            ePhase := E_DL_LoadPortPhase.eLpErr;      // 进故障相 / enter error
            eErr := E_DL_LoadPortErr.eLpErrTmo;       // 故障级：握手超时（与开门超时共用，反证句：输出同为收拢+故障级）/ fault: handshake timeout
        END_IF

    E_DL_LoadPortPhase.eLpMapCmp:
        bDoorOpenCmd := TRUE;                         // 比对：开门保持 / open held
        bDoorCloseCmd := FALSE;                       // 比对：关门撤 / close dropped
        uDiffAcc := 0;                                // 差异计数清零 / difference cleared
        FOR i := DL_LP_SLOT_MIN TO DL_LP_SLOT_MAX DO
            IF aMapExpect[i] <> aMapRead[i] THEN
                uDiffAcc := uDiffAcc + 1;             // 逐位比对差异累加 [片位] / per-slot difference accumulation
            END_IF
        END_FOR
        nMapDiff := uDiffAcc;                         // 差异计数输出 [片位] / difference count output
        IF uDiffAcc = 0 THEN
            bMapMatch := TRUE;                        // 全等：映射一致 / identical: matched
            bReleaseOk := TRUE;                       // 放行许可置位 / release granted
            ePhase := E_DL_LoadPortPhase.eLpRelease;  // 进放行相 / enter release
            eErr := E_DL_LoadPortErr.eLpErrRel;       // 码 0425 / code release
        ELSE
            bMapMatch := FALSE;                       // 不符：映射不一致 / mismatch
            bReleaseOk := FALSE;                      // 不符：拒收 / rejected
            ePhase := E_DL_LoadPortPhase.eLpErr;      // 进故障相（拒收收拢）/ enter error, reject
            eErr := E_DL_LoadPortErr.eLpErrMap;       // 信息级：映射不符（含差异计数）/ info: map mismatch
        END_IF

    E_DL_LoadPortPhase.eLpRelease:
        bDoorOpenCmd := TRUE;                         // 放行：开门保持（取片）/ open held for pick
        bDoorCloseCmd := FALSE;                       // 放行：关门撤 / close dropped
        bReleaseOk := TRUE;                           // 放行许可保持 / release held
        bMapMatch := TRUE;                            // 映射一致保持 / match held
        eErr := E_DL_LoadPortErr.eLpErrRel;           // 码 0425 / code release
        ePhase := E_DL_LoadPortPhase.eLpDone;          // 放行完成进完成相 / release done, enter done

    E_DL_LoadPortPhase.eLpDone:
        bDoorOpenCmd := FALSE;                        // 完成：开门撤 / open dropped
        bDoorCloseCmd := TRUE;                        // 完成：关门收拢 / close for safe collapse
        bReleaseOk := FALSE;                          // 完成：放行撤（本循环结束）/ release dropped
        eErr := E_DL_LoadPortErr.eLpErrRel;           // 码 0425（完成态沿用放行码）/ code release held

    E_DL_LoadPortPhase.eLpErr:
        bDoorOpenCmd := FALSE;                        // 故障相：开门撤 / open dropped
        bDoorCloseCmd := TRUE;                        // 故障相：关门安全收拢 / close for safe collapse
        bReleaseOk := FALSE;                          // 故障相：放行撤 / release dropped
        bMapMatch := FALSE;                           // 故障相：一致标志撤 / match dropped

    ELSE
        ePhase := E_DL_LoadPortPhase.eLpErr;          // 非法相兜底 / illegal-phase fallback
        bDoorOpenCmd := FALSE;                        // 安全态：开门撤 / open dropped, safe side
        bDoorCloseCmd := TRUE;                        // 安全态：关门收拢 / close for safe collapse
        bReleaseOk := FALSE;                          // 安全态：放行撤 / release dropped
        bMapMatch := FALSE;                           // 安全态：一致标志撤 / match dropped
        eErr := E_DL_LoadPortErr.eLpErrTmo;           // 兜底码（超时段，反证句：输出同为收拢+撤放行）/ fallback code

END_CASE
END_FUNCTION_BLOCK

(* ---- FB_DL_LoopAuditTrailWindow.st ---- *)
(*==============================================================================
 * 组件名称 (Component)  : FB_DL_LoopAuditTrailWindow
 * 所属子库 (Sublibrary) : DL_Process
 * 当前版本 (Version)    : 1.0.0
 * 兼容性 (Platform)     : CODESYS 3.5+ / TwinCAT 3 / 汇川 InoProShop / 施耐德 Machine Expert
 *                         仅依赖 Standard.library（R_TRIG / ABS），零厂商私有库
 * 功能描述 (Function)   : 回路整定审计时间窗与变更留痕。维护窗电平内、双人
 *                         确认位同时成立时变更申请放行并留痕（计数 + 锁存）；
 *                         单人确认或窗外申请一律拒绝（独立成因分码 R190），
 *                         窗外申请计数另记审计。与 RecipeManager（参数快照）
 *                         分工：本件管维护窗内变更留痕与双人确认位，是审计
 *                         生命周期管理。
 * 来源标签 (Origin)     : ROADMAP §16.6 R11 池（L736），自研 clean-room
 * 边界语义 (Boundary)   : ① 双人确认 = 双确认位同拍同时电平（单确认位申请
 *                         拒绝成因 eOneOp 独立成员）；
 *                         ② 窗外申请不锁存故障（业务拒绝态），计数 nOutsideCnt
 *                         供审计；
 *                         ③ 留痕锁存 bTrailLatch 至复位沿（审计资产不随窗
 *                         关闭消失）；
 *                         ④ 纯布尔/整型域，无浮点量。
 * 输出语义 (Fallback)   : 【R191】bEnable = FALSE → 放行出口 FALSE（审计放行
 *                         失能必须收敛）；eFault 相 → 放行 FALSE + bError。
 * 码位     (Codes)      : 按 R297 范式零 16# 码位硬编码；错误出口 BOOL+ENUM(eCause)。
 * 红线自检 (Redline)    : 7 项红线已自检：R1 零全局 ✓｜R2 零物理地址 ✓｜R3 纯 IEC ✓
 *                         R4 无浮点域/计数有界 ✓｜R5 双语同行注释 ✓
 *                         R6 CASE 带 ELSE 兜底迁 eFault ✓｜R7 R_TRIG 段 0 无条件刷新 ✓
 * 验收向量 (Acceptance) : V1 窗内 + 双确认 + 申请沿 → bChangeAllow 单拍 +
 *                         nChangeCnt+1 + bTrailLatch=TRUE；
 *                         V2 窗内仅确认位 1 → 拒绝，eDeny=eOneOp；
 *                         V3 窗外申请沿 → 拒绝，eDeny=eOutOfWin，
 *                         nOutsideCnt+1。
 * 修订历史 (Revision)   : 2026-11-20  v1.0.0  R51 首版（批 2 · 序号 9）
 *==============================================================================*)
TYPE E_DL_LawDeny :
(
    eNone     := 0,                          (* 无拒绝（已放行或无申请） / No deny *)
    eOutOfWin := 1,                          (* 窗外申请拒绝 / Outside window *)
    eOneOp    := 2                           (* 单人确认拒绝 / Single-operator deny *)
);
END_TYPE

TYPE E_DL_LawState :
(
    eIdle  := 0,                             (* 待使能 / Idle *)
    eAudit := 10,                            (* 审计判定运行 / Audit run *)
    eFault := 90                             (* 故障锁存相 / Fault latched phase *)
);
END_TYPE

TYPE E_DL_LawCause :
(
    eNone     := 0,                          (* 无故障成因 / No cause *)
    ePhaseBad := 3                           (* 非法相位兜底 / Illegal phase fallback *)
);
END_TYPE

FUNCTION_BLOCK FB_DL_LoopAuditTrailWindow
VAR_INPUT
    bInAuditWin : BOOL := FALSE;             (* 维护窗电平（上层窗判定供给）[-] / Audit-window level *)
    bChangeReq  : BOOL := FALSE;             (* 变更申请电平（上升沿判）[-] / Change request *)
    bConfirmOp1 : BOOL := FALSE;             (* 操作员 1 确认位电平 [-] / Operator 1 confirm *)
    bConfirmOp2 : BOOL := FALSE;             (* 操作员 2 确认位电平 [-] / Operator 2 confirm *)
    bEnable     : BOOL := TRUE;              (* 使能 [-] / Enable *)
    bReset      : BOOL := FALSE;             (* 复位命令，上升沿清全部（含留痕锁存与计数）[-] / Reset command *)
END_VAR
VAR_OUTPUT
    bChangeAllow : BOOL;                     (* 变更放行单拍位 [-] / Change-allow pulse *)
    eDeny        : E_DL_LawDeny;             (* 拒绝成因（信息级逐拍重算，R189） / Deny cause *)
    bTrailLatch  : BOOL;                     (* 窗内变更已留痕锁存（复位沿清，R152） / Trail latch *)
    nChangeCnt   : UDINT;                    (* 窗内变更留痕计数 [次] / In-window change count *)
    nOutsideCnt  : UDINT;                    (* 窗外申请计数（审计）[次] / Outside request count *)
    nDenyCnt     : UDINT;                    (* 拒绝总计数（审计）[次] / Deny count *)
    eState       : E_DL_LawState;            (* 状态出口 / State outlet *)
    eCause       : E_DL_LawCause;            (* 故障成因出口 / Fault cause outlet *)
    bError       : BOOL;                     (* 故障锁存标志 [-] / Fault latch flag *)
END_VAR
VAR
    _eState    : E_DL_LawState := E_DL_LawState.eIdle;     (* 内部相位（CASE 唯一写入目标） / Internal phase *)
    _eCause    : E_DL_LawCause := E_DL_LawCause.eNone;     (* 故障成因锁存量 / Latched cause *)
    rtReq      : R_TRIG;                     (* 申请沿实例，段 0 无条件调用 / Request edge instance *)
    rtReset    : R_TRIG;                     (* 复位沿实例，段 0 无条件调用 / Reset edge instance *)
    _nInWin    : UDINT;                      (* 窗内变更计数锁存 [次] / In-window count latch *)
    _nOutside  : UDINT;                      (* 窗外申请计数锁存 [次] / Outside count latch *)
    _nDeny     : UDINT;                      (* 拒绝计数锁存 [次] / Deny count latch *)
    _bTrail    : BOOL;                       (* 留痕锁存量 [-] / Trail latch work *)
    _bAllow    : BOOL;                       (* 放行单拍量 [-] / Allow pulse work *)
    _bFault    : BOOL;                       (* 故障锁存位 / Latched fault bit *)
END_VAR

(* —— 段 0：沿实例无条件刷新（R228A；纯布尔/整型域无浮点组态闸） —— *)
rtReq(CLK := bChangeReq);                    (* 申请沿每拍必调 / Request edge every scan *)
rtReset(CLK := bReset);                      (* 复位沿每拍必调 / Reset edge every scan *)

(* —— 段 1：单拍量预清零（R107） —— *)
_bAllow := FALSE;                            (* 放行脉冲预清，唯一分支置位 / Allow preset *)
bChangeAllow := FALSE;                       (* 放行出口预清 / Allow outlet preset *)
eDeny := E_DL_LawDeny.eNone;                 (* 拒绝成因预清（信息级逐拍重算） / Deny preset *)

(* —— 段 2：复位沿处理（作用域：清故障 + 清留痕锁存 + 清三计数 + 迁 eIdle，R283 逐项声明） —— *)
IF rtReset.Q THEN
    _bFault := FALSE;                        (* 清故障锁存 / Clear fault *)
    _eCause := E_DL_LawCause.eNone;          (* 清成因 / Clear cause *)
    _bTrail := FALSE;                        (* 清留痕锁存 / Clear trail latch *)
    bTrailLatch := FALSE;                    (* 清留痕出口 / Clear trail outlet *)
    _nInWin := 0;                            (* 清窗内计数 / Clear in-window count *)
    _nOutside := 0;                          (* 清窗外计数 / Clear outside count *)
    _nDeny := 0;                             (* 清拒绝计数 / Clear deny count *)
    _eState := E_DL_LawState.eIdle;          (* 迁待机相 / Back to idle *)
END_IF

(* —— 段 4：CASE 主状态机（ELSE 兜底迁 eFault，红线 6） —— *)
CASE _eState OF
    E_DL_LawState.eIdle:                     (* 待机相 / Idle *)
        IF bEnable AND NOT _bFault THEN
            _eState := E_DL_LawState.eAudit; (* 进入审计 / Enter audit *)
        END_IF
    E_DL_LawState.eAudit:                    (* 审计相：申请沿三分支判定 / Audit *)
        IF NOT bEnable THEN
            _eState := E_DL_LawState.eIdle;  (* 失能回待机 / Back to idle *)
        ELSIF rtReq.Q THEN                   (* 申请沿判定 / On request edge *)
            IF NOT bInAuditWin THEN
                eDeny := E_DL_LawDeny.eOutOfWin;   (* 成因：窗外（独立成员，R190） / Cause: outside *)
                _nOutside := _nOutside + 1;      (* 窗外计数（UDINT 回绕工程安全） / Count outside *)
                _nDeny := _nDeny + 1;            (* 拒绝总计数 / Count deny *)
            ELSIF NOT (bConfirmOp1 AND bConfirmOp2) THEN   (* 双人确认闸（同拍同时电平，边界①） / Two-operator gate *)
                eDeny := E_DL_LawDeny.eOneOp;    (* 成因：单人（独立成员，R190） / Cause: single op *)
                _nDeny := _nDeny + 1;            (* 拒绝总计数 / Count deny *)
            ELSE
                _bAllow := TRUE;             (* 放行单拍 / Allow pulse *)
                _nInWin := _nInWin + 1;      (* 留痕计数 / Count change *)
                _bTrail := TRUE;             (* 留痕锁存置位（复位沿清，边界③） / Set trail latch *)
            END_IF
        END_IF
    E_DL_LawState.eFault:                    (* 故障相：冻结保持，仅复位沿出 / Fault *)
        ;                                    (* 锁存回放（R28） / Replay from latch *)
    ELSE                                     (* 非法相位兜底迁安全态 / Illegal phase fallback *)
        _eState := E_DL_LawState.eFault;     (* 迁故障相 / To fault *)
        _bFault := TRUE;                     (* 同步锁存 / Latch *)
        _eCause := E_DL_LawCause.ePhaseBad;  (* 成因：非法相位 / Cause: illegal phase *)
END_CASE

(* —— 段 5：出口映射（bError/eState 同源，R191） —— *)
bChangeAllow := _bAllow;                     (* 放行脉冲出口 / Allow outlet *)
bTrailLatch := _bTrail;                      (* 留痕锁存出口 / Trail outlet *)
nChangeCnt := _nInWin;                       (* 窗内计数出口 / In-window outlet *)
nOutsideCnt := _nOutside;                    (* 窗外计数出口 / Outside outlet *)
nDenyCnt := _nDeny;                          (* 拒绝计数出口 / Deny outlet *)
bError := _bFault;                           (* 故障标志镜像 / Fault flag mirror *)
eState := _eState;                           (* 状态出口 / State outlet *)
eCause := _eCause;                           (* 成因出口 / Cause outlet *)
END_FUNCTION_BLOCK

(* ---- FB_DL_LotGenealogyLink.st ---- *)
(*
  ==================================================================
  组件名 Component  : FB_DL_LotGenealogyLink
  分类   Category   : DL_Process
  复杂度 Complexity  : 中
  版本   Version    : 1.0.0
  功能   Purpose    : 批次谱系链接（ISA-88 批次谱系公开模型）。64 槽注册表：
                      登记批次（bRegReq）→ 建父子链（bLinkReq，环检测 + 深度
                      上限 16）→ 解链（bUnlinkReq）；nDepth 实时输出 nLotId
                      批次谱系深度；拒绝类结果 bRefused 单脉冲并区分成因
                      bCycleDetected / bDepthExceeded。与
                      FB_DL_TrackBarcodeTrace 单件追踪分工。
  来源   Source     : T2-8-isa-88（ISA-88 批次谱系公开模型）
  溯源   Origin     : ISA-88 批次父子谱系为公开模型语义，clean-room 自研实
                      现，未复制任何厂商私有库源码。
  平台   Platform   : 纯 IEC 61131-3，CODESYS / TwinCAT / InoProShop 通用
  分工声明 Split     : 与 FB_DL_TrackBarcodeTrace 分工——后者做单件条码追踪，
                      本件做批次级父子谱系链维护。
  作者   Author     : 道莅代码库 · PLC 编程专家（R59）
  ------------------------------------------------------------------
  边界 Boundary     :
                      一 操作闸：登记重号 / 注册表满 / 链接任一批次未登记 /
                         解链批次未登记 → bRefused 单脉冲（信息级拒绝，非故
                         障）；环检出 bCycleDetected / 深度超限 bDepthExceeded
                         为独立成因独立标志（R190）；
                      二 深度上限 16：链上行遍历以深度限为界（兼作有界环终
                         止条件），超限拒绝建链；
                      三 环检测：从父批沿父链上行，命中子批即判环，拒绝；
                      四 bLinked / bRefused / bCycleDetected / bDepthExceeded
                         均单拍脉冲，每拍前置清零（纪律③）；
                      五 无除法无浮点（纯整数与数组操作，无除零风险）；无全
                         局变量、无外部变量声明、无物理地址寻址。
  修订记录 Revision  :
    2026-11-21  v1.0.0  R59 首版（批 4 · 序号 20）
  ==================================================================
*)

FUNCTION_BLOCK FB_DL_LotGenealogyLink
VAR_INPUT
    nLotId       : DINT := 0;  // 操作批次号（登记 / 链接子批 / 解链对象）[-] / the operated lot id
    nParentLotId : DINT := 0;  // 父批次号（bLinkReq 方向使用）[-] / the parent lot id
    bRegReq      : BOOL := FALSE; // 登记请求，上升沿生效 [-] / the register request, rising edge
    bLinkReq     : BOOL := FALSE; // 建链请求（nLotId 挂 nParentLotId 下），上升沿生效 [-] / the link request, rising edge
    bUnlinkReq   : BOOL := FALSE; // 解链请求，上升沿生效 [-] / the unlink request, rising edge
END_VAR
VAR_OUTPUT
    bLinked        : BOOL := FALSE; // 建链成功单脉冲（单拍）[-] / the linked one shot pulse
    bRefused       : BOOL := FALSE; // 操作拒绝单脉冲（单拍，成因见独立标志）[-] / the refused one shot pulse
    bCycleDetected : BOOL := FALSE; // 环检出单脉冲（单拍，独立成因）[-] / the cycle detected pulse
    bDepthExceeded : BOOL := FALSE; // 深度超限单脉冲（单拍，独立成因）[-] / the depth exceeded pulse
    nDepth         : INT  := 0;   // nLotId 批次当前谱系深度（根 = 0）[层] / the current depth of the operated lot, the root is zero
    nLinkCnt       : DINT := 0;   // 在册建链总数 [条] / the total link count
    nUsedCnt       : DINT := 0;   // 注册表已用槽数 [槽] / the used slot count
END_VAR
VAR CONSTANT
    DL_LGL_SLOTS  : DINT := 64; // 注册表槽数 [槽] / the registry slot count
    DL_LGL_DEPTH  : INT  := 16; // 谱系深度上限 [层]（兼作上行遍历环界）/ the depth bound, also the walk loop bound
END_VAR
VAR
    aLotId    : ARRAY[0..63] OF DINT; // 批次号槽组（0 = 空槽）/ the lot id slots, zero means empty
    aParentIx : ARRAY[0..63] OF DINT; // 父槽索引组（-1 = 无父）/ the parent slot indexes, minus one means no parent
    rtReg     : R_TRIG; // 登记沿，段 0 无条件刷新 / the register edge
    rtLink    : R_TRIG; // 建链沿，段 0 无条件刷新 / the link edge
    rtUnlink  : R_TRIG; // 解链沿，段 0 无条件刷新 / the unlink edge
    _nI       : DINT;  // 槽遍历索引 / the slot loop index
    _nChild   : DINT;  // 子批槽索引工作量 [槽] / the child slot work index
    _nParent  : DINT;  // 父批槽索引工作量 [槽] / the parent slot work index
    _nWalk    : DINT;  // 上行遍历槽索引 [槽] / the walk slot index
    _nDepth   : INT;   // 深度工作量 [层] / the depth work value
    _nFree    : DINT;  // 空槽索引工作量（-1 = 满）/ the free slot index, minus one means full
    _bFound   : BOOL;  // 槽查找命中工作量 [-] / the slot found work flag
END_VAR

// 段 0｜沿检测无条件周期刷新（禁入分支，R7）/ segment 0, the unconditional refresh
rtReg(CLK := bRegReq); // 登记沿 / the register edge
rtLink(CLK := bLinkReq); // 建链沿 / the link edge
rtUnlink(CLK := bUnlinkReq); // 解链沿 / the unlink edge

// 段 1｜单拍脉冲前置清零（边界四，纪律③）/ segment 1, the per scan pulse preset
bLinked := FALSE; // 建链脉冲预清零 / preset the linked false
bRefused := FALSE; // 拒绝脉冲预清零 / preset the refused false
bCycleDetected := FALSE; // 环脉冲预清零 / preset the cycle false
bDepthExceeded := FALSE; // 深度脉冲预清零 / preset the depth false

// 段 2｜登记操作（重号拒 / 表满拒，边界一）/ segment 2, the register operation
IF rtReg.Q THEN // 登记沿 / the register edge
    IF nLotId <> 0 THEN // 零号保留为空槽哨兵，禁登记 / the zero id reserved, refused
        _bFound := FALSE; // 重号查找清 / clear the dup search
        _nFree := -1; // 空槽查找清（-1 = 满）/ clear the free search
        FOR _nI := 0 TO DL_LGL_SLOTS - 1 DO // 全槽扫描 / per slot
            IF aLotId[_nI] = nLotId THEN // 重号命中 / a dup hit
                _bFound := TRUE; // 记重号 / mark the dup
            ELSIF aLotId[_nI] = 0 THEN // 空槽捕获（记首个）/ capture the first free slot
                IF _nFree < 0 THEN // 尚未捕获 / not captured yet
                    _nFree := _nI; // 记空槽 / mark the free slot
                END_IF
            END_IF
        END_FOR
        IF _bFound OR (_nFree < 0) THEN // 重号或表满拒绝（信息级）/ a dup or full, refused
            bRefused := TRUE; // 置拒绝脉冲 / raise the refused pulse
        ELSE // 受理登记 / accept the registration
            aLotId[_nFree] := nLotId; // 批次号入槽 / store the lot id
            aParentIx[_nFree] := -1; // 无父起步 / start without a parent
            nUsedCnt := nUsedCnt + 1; // 用槽计数推进 / advance the used count
        END_IF
    ELSE // 零号登记拒绝 / the zero id refused
        bRefused := TRUE; // 置拒绝脉冲 / raise the refused pulse
    END_IF
END_IF

// 段 3｜槽定位公共步（子批与父批索引查找）/ segment 3, the slot locating common step
_nChild := -1; // 子批索引清（-1 = 未登记）/ clear the child index
_nParent := -1; // 父批索引清 / clear the parent index
FOR _nI := 0 TO DL_LGL_SLOTS - 1 DO // 全槽查找 / per slot search
    IF aLotId[_nI] = nLotId THEN // 子批命中 / the child hit
        _nChild := _nI; // 记子批槽 / mark the child slot
    END_IF
    IF aLotId[_nI] = nParentLotId THEN // 父批命中 / the parent hit
        _nParent := _nI; // 记父批槽 / mark the parent slot
    END_IF
END_FOR

// 段 4｜谱系深度实时计算（上行遍历以深度限为界，边界二）/ segment 4, the live depth calculation
nDepth := 0; // 深度预置根零 / preset the root zero
IF _nChild >= 0 THEN // 批次在册才算深度 / the depth only for a registered lot
    _nDepth := 0; // 深度清零 / clear the depth
    _nWalk := aParentIx[_nChild]; // 从父槽上行 / walk up from the parent slot
    WHILE (_nWalk >= 0) AND (_nDepth < DL_LGL_DEPTH) DO // 有界上行环 / the bounded walk
        _nDepth := _nDepth + 1; // 深度推进 / advance the depth
        _nWalk := aParentIx[_nWalk]; // 继续上行 / keep walking
    END_WHILE
    nDepth := _nDepth; // 深度出口（超限截断口径）/ the depth outlet, truncated by the bound
END_IF

// 段 5｜建链操作（未登记拒 / 环拒 / 深度超限拒，边界一二三）/ segment 5, the link operation
IF rtLink.Q THEN // 建链沿 / the link edge
    IF (_nChild < 0) OR (_nParent < 0) THEN // 任一批次未登记拒绝 / either unregistered, refused
        bRefused := TRUE; // 置拒绝脉冲 / raise the refused pulse
    ELSE // 双批在册，环与深度闸 / both registered, the cycle and depth gates
        _bFound := FALSE; // 环检出工作量清 / clear the cycle search
        _nDepth := 0; // 深度工作量清 / clear the depth
        _nWalk := _nParent; // 从父批上行 / walk up from the parent
        WHILE (_nWalk >= 0) AND (_nDepth < DL_LGL_DEPTH) DO // 有界上行（深度限兼环界）/ the bounded walk
            IF _nWalk = _nChild THEN // 上行命中子批：环 / the child hit, a cycle
                _bFound := TRUE; // 记环 / mark the cycle
                _nWalk := -1; // 终止遍历 / stop the walk
            ELSE // 未命中继续上行 / not hit, keep walking
                _nWalk := aParentIx[_nWalk]; // 上行一步 / walk one step
                _nDepth := _nDepth + 1; // 深度推进 / advance the depth
            END_IF
        END_WHILE // 环上行结束（R59 修：原误写 END_FOR，编译阻断）/ end of the bounded walk
        IF _bFound THEN // 环检出：拒绝建链（独立成因，R190）/ a cycle detected, refused
            bCycleDetected := TRUE; // 置环脉冲 / raise the cycle pulse
            bRefused := TRUE; // 同步置拒绝脉冲 / raise the refused pulse
        ELSIF (nDepth + 1) > DL_LGL_DEPTH THEN // 子批挂后深度超限：拒绝（独立成因）/ the depth beyond the bound, refused
            bDepthExceeded := TRUE; // 置深度脉冲 / raise the depth pulse
            bRefused := TRUE; // 同步置拒绝脉冲 / raise the refused pulse
        ELSE // 受理建链 / accept the link
            aParentIx[_nChild] := _nParent; // 写父槽索引 / write the parent index
            nLinkCnt := nLinkCnt + 1; // 建链计数推进 / advance the link count
            bLinked := TRUE; // 置建链成功脉冲 / raise the linked pulse
        END_IF
    END_IF
END_IF

// 段 6｜解链操作（未登记拒，成功不脉冲只更新）/ segment 6, the unlink operation
IF rtUnlink.Q THEN // 解链沿 / the unlink edge
    IF _nChild < 0 THEN // 批次未登记拒绝 / unregistered, refused
        bRefused := TRUE; // 置拒绝脉冲 / raise the refused pulse
    ELSIF aParentIx[_nChild] >= 0 THEN // 有父可解 / a parent exists
        aParentIx[_nChild] := -1; // 清父索引 / clear the parent index
        nLinkCnt := nLinkCnt - 1; // 建链计数回落 / drop the link count
        IF nLinkCnt < 0 THEN // 计数防御兜底（不可达分支）/ the unreachable fallback
            nLinkCnt := 0; // 夹回零 / clamp to zero
        END_IF
    END_IF
END_IF
END_FUNCTION_BLOCK

(* ---- FB_DL_LotMergeGate.st ---- *)
(*
  ==================================================================
  组件名 Component  : FB_DL_LotMergeGate
  分类   Category   : DL_Process
  前缀   Naming     : FB_DL_ ｜ b/n/u/f/t/e 类型前缀制（R265）
  版本   Version    : 1.0.1
  功能   Purpose    : 批次合批闸：按「批次数 nLotsReq / 总量 uQtyReq」双门槛
                      收集来料批次，门槛任一满足即转就绪；就绪后 bRelease
                      放行（bReleased=TRUE），放行态可经 bRecall 回迁召回态
                      再放行（合规重入）。配置非法（nLotsReq=0 或 uQtyReq=0）
                      锁存 eFault；累计器溢出钳位 + 信息码，不静默吞量。
                      bResetCmd 上升沿复位同步清账（锁存/累计/状态全清）。
  来源   Source     : t2-8-isa88（ISA-88 批次相语义：借「合批/放行/召回」相
                      命名组织方式，实现零源码复制）
  互引   Cross-ref  : FB_DL_ReworkLotGate（同族批次门禁件：返工拦截闸，本件
                      为合批闸，二者可级联——先返工门禁后合批）；FB_DL_LotGenealogyLink
                      （下游批次谱系链接件，可把本件 eState 变迁喂给它建档）
  平台   Platform   : 纯 IEC 61131-3（R_TRIG/ENUM+CASE/UDINT 四则）
  依赖   Depends    : 仅 Standard.library（R_TRIG 属标准件）
  归属   Ownership  : E_DL_MergeState 属主为本文件（全库唯一定义，R264）；
                      引用件只引用不重声明。
  红线   Redline    : R1 零全局/VAR_EXTERNAL/R2 零 %I/%Q/R3 纯 IEC 标准
                      R4 无浮点（纯整数与布尔，无除法面）/R5 全变量双语同行
                      注释/R6 ENUM+CASE 含 ELSE 兜底，eFault 分支显式出现
                      R7 四个 R_TRIG 段 0 无条件刷新/R8 溢出钳位常量化
  契约   Contract   : bEnable 未设引脚（本件无失能面，复位沿即总闸）；uLotQty
                      在 eIdle 相首个 bLotIn 沿入账、eCollecting 相后续沿逐批
                      累加；bReleased 仅在 eReleased 相为 TRUE（召回/复位即撤）。
  错误码 Codes      : 01【故障级·锁存】配置非法（nLotsReq=0 或 uQtyReq=0），
                      锁存至复位沿
                      02【信息级】累计器溢出钳位（uQtyAcc 饱和于 UDINT 上限）
                      03【故障级·锁存】非法状态拦截（ELSE 兜底）
  码位反证 Note     : 01/02/03 分立依据（R90）：01 在配置面、02 在台账面
                      （功能不受影响，bError 不置）、03 在状态面可观测；
                      02 为信息级不置 bError，与 01/03 故障级双通道可区分。
  验收   Acceptance : V1 3 批门槛收满 → eReady ｜ V2 eReady + bRelease →
                      eReleased + bReleased ｜ V3 eReleased + bRecall →
                      eRecalled + bReleased 撤 ｜ V4 eRecalled + bRelease →
                      eReleased（合规重入）｜ V5 nLotsReq=0 → 锁存 01 ｜
                      V6 溢出钳位 → 码 02（不置 bError）｜ V7 复位沿 → 全清
                      回 eIdle ｜ V8 强改非法态 → ELSE 锁存 03
  变更   Revision   : 2026-11-22  v1.0.0  R66 首版（编码阶段批 4 序 9）
                      2026-11-22  v1.0.1  R67 点修（L3）：删除 eFault 分支
                      死迁出式 IF NOT _bFaultLatch → eIdle（迁入 eFault 必伴
                      锁存，清锁存的复位沿同拍已先行置 eIdle，该式结构性不可
                      达）；eFault 相出口仅保留锁存解除路径（复位沿，段 2）。
                      按「结构性不可达防御统一记账口径」登记：eIdle 相
                      uLotQty > LMG_U_MAX 留档型防御（L2）保留不动（UDINT
                      入口域上不可达，留档备审计）。
  ==================================================================
*)
TYPE E_DL_MergeState :
(
    eIdle      := 0,   // 待机：无收集中批次 / idle, no batch being collected
    eCollecting:= 10,  // 收集中：累计未达任一门槛 / collecting, neither threshold met
    eReady     := 20,  // 就绪：门槛任一满足，待放行 / ready, a threshold met, awaiting release
    eReleased  := 30,  // 放行：bReleased=TRUE，可召回 / released, bReleased true, recallable
    eRecalled  := 40,  // 召回：放行被撤回，可再放行 / recalled, the release withdrawn, re releasable
    eFault     := 50   // 锁存故障：复位沿解除 / the latched fault, released by the reset edge
);
END_TYPE

FUNCTION_BLOCK FB_DL_LotMergeGate
VAR_INPUT
    bLotIn   : BOOL := FALSE;  // 来料批次脉冲（上升沿入账）[-] / the incoming lot pulse, counted on the rising edge
    uLotQty  : UDINT := 0;     // 当前批次数量 [件] / the current lot quantity [pc]
    nLotsReq : UDINT := 0;     // 批次数门槛 [批]，须 ≥ 1（=0 判配置非法）/ the lots threshold, at least one
    uQtyReq  : UDINT := 0;     // 总量门槛 [件]，须 ≥ 1（=0 判配置非法）/ the quantity threshold, at least one
    bRelease : BOOL := FALSE;  // 放行指令（上升沿生效）[-] / the release command, effective on the rising edge
    bRecall  : BOOL := FALSE;  // 召回指令（上升沿生效）[-] / the recall command, effective on the rising edge
    bResetCmd: BOOL := FALSE;  // 复位指令（上升沿同步清账）[-] / the reset command, clears the books on the rising edge
END_VAR
VAR_OUTPUT
    eState   : E_DL_MergeState := E_DL_MergeState.eIdle; // 状态机出口 [状态] / the state machine outlet
    uLotsAcc : UDINT := UDINT#0;   // 已收批次数 [批] / the collected lots count
    uQtyAcc  : UDINT := UDINT#0;   // 已收总量 [件]（溢出钳位于 UDINT 上限）/ the collected quantity, saturated
    bReleased: BOOL := FALSE;      // 放行态指示（仅 eReleased 相为 TRUE）[-] / the released indicator, true only in the released phase
    bError   : BOOL := FALSE;      // 故障锁存标志（复位沿清除，R45 配对）/ the latched fault flag, cleared by the reset edge
    uErrorId : UDINT := 16#0000_0000; // 错误码，0=正常；锁存回放至复位沿 [码] / the error code replayed to the reset edge
END_VAR
VAR
    _eState      : E_DL_MergeState := E_DL_MergeState.eIdle; // 内部状态寄存器 / the internal state register
    _bFaultLatch : BOOL := FALSE;   // 故障锁存副本（仅复位沿清除）/ the fault latch copy, cleared only by the reset edge
    _uLatch      : UDINT := 16#0000_0000; // 故障码锁存副本（FB33-1）/ the latched code copy
    _bQtySat     : BOOL := FALSE;   // 本拍溢出钳位信息位（单拍，段 6 映射）/ the per scan saturation info bit
    rtLotIn      : R_TRIG;          // 来料沿实例，段 0 无条件刷新 / the lot edge instance refreshed unconditionally
    rtRelease    : R_TRIG;          // 放行沿实例，段 0 无条件刷新 / the release edge instance refreshed unconditionally
    rtRecall     : R_TRIG;          // 召回沿实例，段 0 无条件刷新 / the recall edge instance refreshed unconditionally
    rtReset      : R_TRIG;          // 复位沿实例，段 0 无条件刷新（锁存解除可达边）/ the reset edge instance, the reachable release edge
END_VAR
VAR CONSTANT
    LMG_U_MAX    : UDINT := 4294967295;   // UDINT 上限哨兵 [件] / the UDINT ceiling sentinel
    LMG_ERR_NONE : UDINT := 16#0000_0000; // 无错误 [码] / no error [code]
    LMG_ERR_CFG  : UDINT := 16#0000_0001; // 码 01：配置非法（锁存）/ code 01, illegal configuration, latched
    LMG_ERR_SAT  : UDINT := 16#0000_0002; // 码 02：累计器溢出钳位（信息级）/ code 02, accumulator saturation, info level
    LMG_ERR_ILL  : UDINT := 16#0000_0003; // 码 03：非法状态（锁存）/ code 03, illegal state, latched
END_VAR

(*------------------------------------------------------------------------------
 * 段 0｜沿检测无条件刷新区（红线 R7）：严禁移入 IF / CASE
 *      The edge instances refresh unconditionally, never inside a branch
 *-----------------------------------------------------------------------------*)
rtLotIn(CLK := bLotIn);        // 来料沿 / the lot edge
rtRelease(CLK := bRelease);    // 放行沿 / the release edge
rtRecall(CLK := bRecall);      // 召回沿 / the recall edge
rtReset(CLK := bResetCmd);     // 复位沿 / the reset edge

(*------------------------------------------------------------------------------
 * 段 1｜错误码本拍预置 + 信息位复位（当前周期事实）
 *      The error code and the info bit are per scan facts
 *-----------------------------------------------------------------------------*)
uErrorId := LMG_ERR_NONE;      // 预置无错误（锁存值随后回放覆盖）/ preset none, the latch replays over it
_bQtySat := FALSE;             // 单拍信息位复位 / reset the single scan info bit

(*------------------------------------------------------------------------------
 * 段 2｜复位沿：同步清账（锁存/累计/状态/bReleased 全清回 eIdle）
 *      The reset edge clears the books synchronously
 *-----------------------------------------------------------------------------*)
IF rtReset.Q THEN
    _bFaultLatch := FALSE;     // 清锁存副本 / clear the latch copy
    _uLatch := LMG_ERR_NONE;   // 清锁存码 / clear the latched code
    uLotsAcc := UDINT#0;       // 清批次数台账 / clear the lots ledger
    uQtyAcc := UDINT#0;        // 清总量台账 / clear the quantity ledger
    _eState := E_DL_MergeState.eIdle;  // 回待机相 / back to idle
    bReleased := FALSE;        // 撤放行指示 / withdraw the release indicator
END_IF

(*------------------------------------------------------------------------------
 * 段 3｜配置闸（锁存归因，成因独立 R190）：门槛任一为 0 即锁存 eFault
 *      The configuration gate, either threshold of zero latches the fault
 *-----------------------------------------------------------------------------*)
IF (nLotsReq = UDINT#0) OR (uQtyReq = UDINT#0) THEN
    _bFaultLatch := TRUE;      // 锁存置位 / latch on
    _uLatch := LMG_ERR_CFG;    // 配置非法码 / the configuration code
END_IF

(*------------------------------------------------------------------------------
 * 段 4｜状态机（ENUM + CASE，含 ELSE 兜底；eFault 分支显式出现）
 *      本拍合法事件优先于故障推断（R275 同拍竞态）：复位沿已先行消化
 *      The state machine, legal events first, the reset edge already consumed above
 *-----------------------------------------------------------------------------*)
IF _bFaultLatch THEN
    _eState := E_DL_MergeState.eFault;   // 锁存强制故障相 / the latch forces the fault phase
END_IF
CASE _eState OF
E_DL_MergeState.eIdle:                   // 待机相 / the idle phase
    IF rtLotIn.Q THEN                    // 首批入账 / the first lot books in
        uLotsAcc := UDINT#1;             // 批次计数起账 / start the lots ledger
        IF uLotQty > LMG_U_MAX THEN      // 批量溢出闸（结构性不可达，留档）/ the per lot overflow gate
            uQtyAcc := LMG_U_MAX;        // 钳上限 / clamp to the ceiling
            _bQtySat := TRUE;            // 记信息位 / mark the info bit
        ELSE
            uQtyAcc := uLotQty;          // 总量入账 / book the quantity
        END_IF
        IF (uLotsAcc >= nLotsReq) OR (uQtyAcc >= uQtyReq) THEN
            _eState := E_DL_MergeState.eReady;   // 门槛即达直接就绪 / ready immediately when a threshold is met
        ELSE
            _eState := E_DL_MergeState.eCollecting;  // 否则迁入收集相 / else enter the collecting phase
        END_IF
    END_IF
E_DL_MergeState.eCollecting:             // 收集相 / the collecting phase
    IF rtLotIn.Q THEN                    // 后续批逐批入账 / each following lot books in
        IF uLotsAcc < LMG_U_MAX THEN     // 批次计数溢出钳位 / the lots count saturation clamp
            uLotsAcc := uLotsAcc + UDINT#1;
        ELSE
            _bQtySat := TRUE;            // 批次计数饱和记信息位 / mark the info bit
        END_IF
        IF uQtyAcc > LMG_U_MAX - uLotQty THEN  // 总量溢出预判（先闸后加，禁回绕）/ the quantity overflow preview, gate before adding
            uQtyAcc := LMG_U_MAX;        // 钳上限 / clamp to the ceiling
            _bQtySat := TRUE;            // 记信息位 / mark the info bit
        ELSE
            uQtyAcc := uQtyAcc + uLotQty;  // 安全累加 / the safe accumulation
        END_IF
        IF (uLotsAcc >= nLotsReq) OR (uQtyAcc >= uQtyReq) THEN
            _eState := E_DL_MergeState.eReady;   // 门槛满足迁就绪 / the threshold met, enter ready
        END_IF
    END_IF
E_DL_MergeState.eReady:                  // 就绪相 / the ready phase
    IF rtRelease.Q THEN                  // 放行沿 / the release edge
        _eState := E_DL_MergeState.eReleased;  // 迁入放行相 / enter the released phase
    END_IF
E_DL_MergeState.eReleased:               // 放行相：驻留相（可召回，非单拍回迁）/ the released phase, dwell by design
    bReleased := TRUE;                   // 放行指示与状态同源（R191 名实双出口）/ the indicator mirrors the state
    IF rtRecall.Q THEN                   // 召回沿 / the recall edge
        _eState := E_DL_MergeState.eRecalled;  // 回迁召回相 / enter the recalled phase
    END_IF
E_DL_MergeState.eRecalled:               // 召回相 / the recalled phase
    bReleased := FALSE;                  // 撤放行指示（名实双出口）/ withdraw the indicator
    IF rtRelease.Q THEN                  // 再放行沿（合规重入，头注 V4）/ the re release edge
        _eState := E_DL_MergeState.eReleased;  // 回迁放行相 / back to the released phase
    END_IF
E_DL_MergeState.eFault:                  // 故障相（显式分支）：锁存驻留，解除仅由复位沿承担
    bReleased := FALSE;                  // 故障相撤放行指示 / withdraw the indicator in the fault phase
    // 失能/故障相串清账：bReleased 已撤；台账 uLotsAcc/uQtyAcc 故意保留供审计
    // 回放（锁存回放原则：不在故障相清账，账面随复位沿统一清，R 锁存回放）
    // the ledgers are deliberately kept for audit replay, cleared by the reset edge
    // v1.0.1：本相无迁出式——锁存解除与 eIdle 回迁由复位沿（段 2）同拍承担，
    // 原 IF NOT _bFaultLatch → eIdle 为结构性不可达死代码，已删（R67 L3）
    // the latch release and the idle return are owned by the reset edge alone
ELSE                                     // 非法状态兜底（R 非法态拦截，不静默）
    _eState := E_DL_MergeState.eFault;   // 强制故障相 / force the fault phase
    _bFaultLatch := TRUE;                // 锁存置位 / latch on
    _uLatch := LMG_ERR_ILL;              // 非法状态码 / the illegal state code
END_CASE

(*------------------------------------------------------------------------------
 * 段 5｜出口映射（名实双出口 R191）：状态/锁存/信息码单点映射
 *      The outlet mapping, the state, the latch and the info code from one point
 *-----------------------------------------------------------------------------*)
IF _bFaultLatch THEN
    bError := TRUE;                      // 故障标志（R45 配对）/ the fault flag
    uErrorId := _uLatch;                 // 锁存回放 / the latched replay
ELSE
    bError := FALSE;                     // 无锁存无故障 / no latch no fault
    IF _bQtySat THEN
        uErrorId := LMG_ERR_SAT;         // 信息级码（不置 bError，功能不受影响）/ the info code, no fault flag
    END_IF
END_IF
IF _eState = E_DL_MergeState.eReleased THEN
    bReleased := TRUE;                   // 放行指示终判（唯一来源） / the release indicator final verdict
ELSE
    bReleased := FALSE;                  // 其余相一律撤 / withdrawn in every other phase
END_IF
eState := _eState;                       // 状态出口 / publish the state
END_FUNCTION_BLOCK

(* ---- FB_DL_LotoSequence.st ---- *)
(*
  ==================================================================
  组件名 Component  : FB_DL_LotoSequence
  分类   Category   : DL_Process
  复杂度 Complexity  : 中
  版本   Version    : 1.0.0
  功能   Purpose    : LOTO 上锁挂牌流程（OSHA 公开流程语义）。能量隔离点逐
                      点确认（8 点上限）+ 挂牌台账确认 → 上锁 eLocked；解锁
                      前试启验证窗：窗内出现运动反馈（bMotionFb）判隔离失效
                      锁存 eFault，窗到期无运动才放行 eUnlocked。与
                      FB_DL_GuardLockDoor 单门互锁分工。
  来源   Source     : self-std（OSHA LOTO 公开流程语义）
  溯源   Origin     : OSHA 1910.147 上锁挂牌公开流程语义，clean-room 自研
                      实现，未复制任何厂商私有库源码。
  平台   Platform   : 纯 IEC 61131-3（Standard.library: TON / R_TRIG，无私有库）
  分工声明 Split     : 与 FB_DL_GuardLockDoor 分工——后者做单门互锁，本件
                      做多能量隔离点 LOTO 流程。
  作者   Author     : 道莅代码库 · PLC 编程专家（R59）
  ------------------------------------------------------------------
  边界 Boundary     :
                      一 安全语义：eFault / eIsolate / eIdle 相 bLocked 强制
                         假（安全侧只有 eLocked / eTryVerify 两相上锁口径）；
                      二 试启验证窗到期即放行（窗口末退出迁移，纪律④）；窗
                         内运动反馈 = 隔离失效（独立成因 bFault，R190）；
                      三 上锁判据 = 全部隔离点确认 AND 挂牌台账完成（双闸缺
                         一不迁相）；
                      四 组态域闸：nIsoCnt ∈ [1..8]，越域锁存 bError（解除
                         = bReset 沿，R188）；故障解除路径 = bReset 沿（唯
                         一路径，R188 声明）；
                      五 定时器与沿检测全部段 0 无条件周期刷新（R7）；
                      六 无全局变量、无外部变量声明、无物理地址寻址。
  修订记录 Revision  :
    2026-11-21  v1.0.0  R59 首版（批 3 · 序号 15）
  ==================================================================
*)

TYPE E_DL_LotoPhase :
(
    eLotoIdle      := 0,  // 空闲：等上锁请求 / idle, awaiting the lock request
    eLotoIsolate   := 10, // 隔离确认：逐点确认与挂牌 / the isolating confirm
    eLotoLocked    := 20, // 已上锁：隔离生效 / the locked state
    eLotoTryVerify := 30, // 解锁前试启验证窗 / the try start verify window
    eLotoUnlocked  := 40, // 已解锁：验证通过放行 / the unlocked state
    eLotoFault     := 90  // 隔离失效锁存：仅复位可清 / the isolation failure latch
);
END_TYPE

FUNCTION_BLOCK FB_DL_LotoSequence
VAR_INPUT
    aIsoCfm    : ARRAY[0..7] OF BOOL; // 隔离点逐点确认组（TRUE = 已隔离确认）[-] / the isolation point confirms
    nIsoCnt    : INT  := 4;      // 隔离点数 [点]，域 1..8 / the isolation point count, one through eight
    bTagLedger : BOOL := FALSE;  // 挂牌台账完成确认 [-] / the tag ledger completed confirm
    bReqLock   : BOOL := FALSE;  // 上锁请求，上升沿生效 [-] / the lock request, rising edge effective
    bReqUnlock : BOOL := FALSE;  // 解锁请求，上升沿生效 [-] / the unlock request, rising edge effective
    bMotionFb  : BOOL := FALSE;  // 试启运动反馈，TRUE = 检测到转动 [-] / the try start motion feedback, true = motion detected
    tTryWin    : TIME := T#10S; // 试启验证窗 [毫秒] / the try start verify window [millisecond]
    bReset     : BOOL := FALSE; // 故障与组态复位，上升沿生效 [-] / the fault and config reset, rising edge
END_VAR
VAR_OUTPUT
    eState     : E_DL_LotoPhase := E_DL_LotoPhase.eLotoIdle; // 流程状态输出 [-] / the process state outlet
    bLocked    : BOOL := FALSE; // 上锁口径输出（eLocked / eTryVerify 两相）[-] / the locked verdict outlet
    bReadyUnlock: BOOL := FALSE; // 解锁放行指示（eUnlocked 相）[-] / the unlock release indicator
    nIsoOkCnt  : INT  := 0;   // 已确认隔离点数 [点] / the confirmed isolation point count
    bFault     : BOOL := FALSE; // 隔离失效故障锁存（解除 = bReset 沿）[-] / the isolation failure latch
    bError     : BOOL := FALSE; // 组态域闸故障锁存 [-] / the config gate fault latch
END_VAR
VAR CONSTANT
    DL_LOTO_ISOMAX : INT := 8; // 隔离点容量上界 [点] / the isolation point capacity bound
END_VAR
VAR
    _ePhase  : E_DL_LotoPhase := E_DL_LotoPhase.eLotoIdle; // 内部相位，CASE 唯一写入目标 / the internal phase, the single CASE write target
    _nOk     : INT := 0;   // 已确认点数工作量 [点] / the confirmed count work value
    _nI      : DINT;       // 隔离点遍历索引 / the isolation point loop index
    _bInit   : BOOL := FALSE; // 首拍初始化标志（R310，真实使用：首拍安全态预置）/ the first scan flag, real use
    rtLock   : R_TRIG;     // 上锁请求沿，段 0 无条件刷新 / the lock request edge
    rtUnlock : R_TRIG;     // 解锁请求沿，段 0 无条件刷新 / the unlock request edge
    rtReset  : R_TRIG;     // 复位沿，段 0 无条件刷新 / the reset edge
    tonTry   : TON;        // 试启验证窗，段 0 无条件刷新 / the try start verify window
END_VAR

// 段 0｜定时器与沿检测无条件周期刷新（禁入分支，R7）/ segment 0, the unconditional refresh
rtLock(CLK := bReqLock); // 上锁沿 / the lock edge
rtUnlock(CLK := bReqUnlock); // 解锁沿 / the unlock edge
rtReset(CLK := bReset); // 复位沿 / the reset edge
tonTry(IN := (_ePhase = E_DL_LotoPhase.eLotoTryVerify), PT := tTryWin); // 试启验证窗 / the verify window

// 段 1｜首拍初始化（R310 真实使用路径）：安全态显式预置 / segment 1, the first scan init, the safe preset
IF NOT _bInit THEN // 首拍一拍 / the first scan
    _bInit := TRUE; // 置首拍标志 / raise the flag
    _ePhase := E_DL_LotoPhase.eLotoIdle; // 相位显式安全预置 / the explicit safe phase preset
END_IF

// 段 2｜组态域闸与复位（边界四，解除路径 = bReset 沿，R188）/ segment 2, the config gate and the reset
IF (nIsoCnt < 1) OR (nIsoCnt > DL_LOTO_ISOMAX) THEN // 点数越域 / the point count out of domain
    bError := TRUE; // 置域闸锁存 / raise the config latch
END_IF
IF rtReset.Q THEN // 复位沿 / the reset edge
    bError := FALSE; // 清域闸锁存 / clear the config latch
    IF _ePhase = E_DL_LotoPhase.eLotoFault THEN // 仅故障相消化复位迁相 / only the fault phase consumes the reset
        _ePhase := E_DL_LotoPhase.eLotoIdle; // 回空闲（解除路径唯一，R188）/ back to idle, the unique release
    END_IF
END_IF

// 段 3｜隔离点确认计数（逐点确认口径）/ segment 3, the isolation confirm count
_nOk := 0; // 计数清零 / clear the count
FOR _nI := 0 TO DL_LOTO_ISOMAX - 1 DO // 逐点遍历 / per point
    IF (_nI < nIsoCnt) AND aIsoCfm[_nI] THEN // 组态界内已确认点 / a confirmed point inside the config bound
        _nOk := _nOk + 1; // 计数推进 / advance the count
    END_IF
END_FOR
nIsoOkCnt := _nOk; // 确认数出口 / the confirm count outlet

// 段 4｜相位机：ENUM + CASE，含 ELSE 非法相位兜底（R6 / R128）/ segment 4, the phase machine
CASE _ePhase OF

E_DL_LotoPhase.eLotoIdle: // 空闲相 / the idle phase
    IF rtLock.Q AND (NOT bError) AND (NOT bFault) THEN // 受理上锁请求（组态合法且无故障）/ accept the lock request
        _ePhase := E_DL_LotoPhase.eLotoIsolate; // 迁隔离确认相 / to the isolate phase
    END_IF

E_DL_LotoPhase.eLotoIsolate: // 隔离确认相 / the isolate phase
    IF bFault THEN // 隔离期间失效（独立成因）/ a failure during the isolation
        _ePhase := E_DL_LotoPhase.eLotoFault; // 迁故障锁存相 / to the fault phase
    ELSIF rtUnlock.Q THEN // 隔离期撤单 / a request withdrawn
        _ePhase := E_DL_LotoPhase.eLotoIdle; // 回空闲 / back to idle
    ELSIF (_nOk >= nIsoCnt) AND bTagLedger AND (NOT bError) THEN // 双闸齐 + 组态合法（R59 修：堵 0 隔离点上锁）/ the dual gates met and the config sane
        _ePhase := E_DL_LotoPhase.eLotoLocked; // 迁上锁相 / to the locked phase
    END_IF

E_DL_LotoPhase.eLotoLocked: // 已上锁相 / the locked phase
    IF bFault THEN // 锁定期失效 / a failure while locked
        _ePhase := E_DL_LotoPhase.eLotoFault; // 迁故障相 / to the fault phase
    ELSIF rtUnlock.Q THEN // 受理解锁请求进验证窗 / accept the unlock into the verify window
        _ePhase := E_DL_LotoPhase.eLotoTryVerify; // 迁试启验证相 / to the try verify phase
    END_IF

E_DL_LotoPhase.eLotoTryVerify: // 试启验证相（窗口末退出迁移，边界二）/ the try verify phase
    IF bMotionFb THEN // 窗内检测到转动：隔离失效（独立成因，R190）/ a motion detected, the isolation failure
        _ePhase := E_DL_LotoPhase.eLotoFault; // 迁故障锁存相 / to the fault phase
    ELSIF tonTry.Q THEN // 验证窗到期无运动：放行（窗口末退出迁移）/ the window expired without motion, release
        _ePhase := E_DL_LotoPhase.eLotoUnlocked; // 迁已解锁相 / to the unlocked phase
    END_IF

E_DL_LotoPhase.eLotoUnlocked: // 已解锁相 / the unlocked phase
    IF bFault THEN // 解锁态失效 / a failure while unlocked
        _ePhase := E_DL_LotoPhase.eLotoFault; // 迁故障相 / to the fault phase
    ELSIF rtLock.Q AND (NOT bError) THEN // 重新上锁请求 / a new lock request
        _ePhase := E_DL_LotoPhase.eLotoIsolate; // 迁隔离确认相 / to the isolate phase
    END_IF

E_DL_LotoPhase.eLotoFault: // 故障锁存相：仅复位可清（迁相由段 2 复位分支消化，本相驻留无动作）/ the fault latch phase, the migrate in the reset branch

ELSE // 非法相位兜底（R128）/ the illegal phase fallback
    _ePhase := E_DL_LotoPhase.eLotoIdle; // 回空闲安全相 / back to the safe idle
END_CASE

// 段 5｜统一出口（边界一安全口径）/ segment 5, the unified outlet
bLocked := (_ePhase = E_DL_LotoPhase.eLotoLocked) OR (_ePhase = E_DL_LotoPhase.eLotoTryVerify); // 上锁口径双相 / the locked dual phases
bReadyUnlock := (_ePhase = E_DL_LotoPhase.eLotoUnlocked); // 放行指示 / the release indicator
bFault := (_ePhase = E_DL_LotoPhase.eLotoFault); // 故障锁存位与相位同源（R191 名实双出口）/ the fault latch shares the phase
eState := _ePhase; // 状态出口 / the state outlet
END_FUNCTION_BLOCK

(* ---- FB_DL_LyoPressureRiseTestSeq.st ---- *)
(*
  Name: FB_DL_LyoPressureRiseTestSeq
  Category: DL_Process
  Version: 1.0.0
  Round: R91 / 2026-11-25
  开源溯源：clean-room 自研（族 制药冻干真空冷冻干燥，ST 开源生态实测 0 命中，无外部代码引入）
  功能：1) 压力升测试序状态机，七相推进：待机 → 隔离 → 稳压 → 计时 → 判定 → 复压 → 完成。
           待机相等 xStart 上升沿且腔体已达起始真空度（否则只置信息级码 0221 不放行）；
           隔离相关隔离阀并等阀关到位反馈；稳压相等压力稳定 tSettleS（消除吸附气体影响）；
           计时相记录起点压力并等 tTestS；判定相算泄漏率 Q = dP * V / t 并判定；
           复压相开通气阀复压并等 tRepressS，完成相置 xDone 并保持到撤令。
        2) 泄漏超限中止：判定相算得 Q > fLeakMaxMbarLs 即判不合格并锁码 0229、进故障相，
           同时撤销全部阀门命令（安全侧：通气阀关、隔离阀保持关闭，防误开腔）。
        3) 每相独立超时 + 整序总超时：相定时器给正常推进点，相超时定时器给「定时 + 裕量」越限点，
           tonTotal 兜底整序总时长，四者并发监视，任一命中立即锁码进故障相。
  边界条件：1) 非有限值闸：压力、容积、泄漏上限先过 NOT(x > -DL_BIG AND x < DL_BIG)，同时拦 NaN 与 Inf；
           命中即锁码 0228 进故障相，绝不把 NaN 拿去与真空度阈值比较（NaN 比较恒假会伪装成「已达真空」，R19）。
        2) 时间参数零闸：tSettleS / tTestS / tRepressS <= T#0S 时对应相定时器立即置 Q（等价跳过该相），
           属合法调试组态；但计时相零时长会计得 Q = 0/0，故在判定相入口对实际计时 > DL_EPS 做显式零闸，
           零闸不通过即锁码 0224 而非输出无穷大泄漏率。
        3) 容积零闸：fVolumeL <= DL_EPS 时泄漏率不可算（乘子为零会把「未组态」伪装成「密封完好」），
           在判定相锁码 0228 并判不合格。
        4) 压力方向：升压为负（隔离后压力下降）说明隔离阀未关严或泵未停，判不合格锁码 0229，
           不取绝对值掩盖隔离失效。
        5) 定时器周期刷新（R7）：十个 TON 与复位边沿全部在 CASE 之外无条件调用。
        6) 故障解除路径：故障相内 xReset 上升沿 AND NOT xFault AND 入参有限 → 清锁存回待机，
           回待机后必须重新给 xStart 上升沿才能再测（不自恢复）。
        7) 状态机兜底：CASE 全态覆盖 + ELSE 强制回故障相并置码 0230、清全部输出。
  量纲自证：Q = dP [mbar] * V [L] / t [s] = mbar*L/s，与 fLeakMaxMbarLs 同量纲，可直接比较；
           所有时间引脚为 [TIME]，相超时点 = [TIME] + [TIME] = [TIME]，与 TON 的 PT 同量纲。
  码表 Error codes（本件子带 0091_022x，故障级一律 3 行内置 _uFault/_bFault/_eState）:
    16#0091_0221 信息级：腔体压力未达起始真空度，禁止启动测试（不置故障位）
    16#0091_0222 故障级：隔离相超时（隔离阀未关到位）
    16#0091_0223 故障级：稳压相超时
    16#0091_0224 故障级：计时相超时或实际计时为零（泄漏率不可算）
    16#0091_0225 故障级：复压相超时
    16#0091_0226 故障级：整序总超时
    16#0091_0227 故障级：外部故障输入 xFault
    16#0091_0228 故障级：压力/容积/限值入参非有限或容积未组态
    16#0091_0229 故障级：泄漏率超限（不合格，或升压为负即隔离失效）
    16#0091_0230 故障级：状态机落 ELSE 兜底（非法相位 ID）

  修订历史 Revision :
    2026-11-25  v1.0.0  R91 首版
*)

TYPE E_DL_LyoPrTestState :
(
    eLyoPrIdle    := 0,     // 待机：等启动沿与起始真空度 / Idle, awaiting the start edge and base vacuum
    eLyoPrIsolate := 10,    // 隔离：关隔离阀等到位反馈 / Isolate, closing the isolation valve
    eLyoPrSettle  := 20,    // 稳压：等吸附气体平衡 / Settle, awaiting desorption equilibrium
    eLyoPrTiming  := 30,    // 计时：记录起点压力并等测试窗 / Timing, base pressure captured
    eLyoPrJudge   := 40,    // 判定：算泄漏率并判合格 / Judge, computing and comparing the leak rate
    eLyoPrRepress := 50,    // 复压：开通气阀复压 / Repressurise, opening the vent valve
    eLyoPrDone    := 60,    // 完成：保持至撤令 / Done, held until the command is released
    eLyoPrFault   := 90     // 故障：锁存待解除 / Fault, latched awaiting release
);
END_TYPE

FUNCTION_BLOCK FB_DL_LyoPressureRiseTestSeq
VAR_INPUT
    xStart           : BOOL;   // 测试启动指令（上升沿有效）[bool] / Test start command, edge triggered [bool]
    xReset           : BOOL;   // 故障复位（上升沿有效）[bool] / Fault reset, rising edge [bool]
    xFault           : BOOL;   // 外部故障汇总 [bool] / External fault aggregate [bool]
    xIsoValveClosedFb : BOOL;  // 隔离阀关到位反馈 [bool] / Isolation valve closed feedback [bool]
    fChamberPressMbar : REAL;  // 腔体实测压力 [mbar] / Measured chamber pressure [mbar]
    fVolumeL         : REAL;   // 腔体（含管路）内容积 [L] / Chamber and piping internal volume [L]
    fLeakMaxMbarLs   : REAL;   // 泄漏率合格上限 [mbar*L/s] / Leak rate acceptance limit [mbar*L/s]
    tSettleS         : TIME;   // 稳压相设定时长 [TIME] / Settle phase duration [TIME]
    tTestS           : TIME;   // 计时相设定时长 [TIME] / Timing phase duration [TIME]
    tRepressS        : TIME;   // 复压相设定时长 [TIME] / Repressurisation phase duration [TIME]
END_VAR
VAR_OUTPUT
    xIsoValveCmd     : BOOL;   // 隔离阀关闭命令（安全侧：故障时保持关闭）[bool] / Isolation valve close command [bool]
    xVentCmd         : BOOL;   // 通气复压阀命令（安全侧：故障时关）[bool] / Vent valve command, fail-safe [bool]
    fLeakRateMbarLs  : REAL;   // 实测泄漏率 [mbar*L/s] / Measured leak rate [mbar*L/s]
    xTestPass        : BOOL;   // 测试合格（保持至撤令）[bool] / Test passed, held until release [bool]
    xDone            : BOOL;   // 测试完成保持位 [bool] / Test complete held flag [bool]
    xBusy            : BOOL;   // 测试进行中 [bool] / Test sequence busy [bool]
    eState           : E_DL_LyoPrTestState;   // 状态出口，段尾单点映射 / State outlet, single-point mapped
    nErrId           : UDINT;  // 事件码，0 = 无事件 / Event code, 0 = none
END_VAR
VAR
    tonIso           : TON;    // 隔离相正常定时 [TIME] / Isolation phase timer
    tonIsoOv         : TON;    // 隔离相超时定时 [TIME] / Isolation phase overrun timer
    tonSettle        : TON;    // 稳压相正常定时 [TIME] / Settle phase timer
    tonSettleOv      : TON;    // 稳压相超时定时 [TIME] / Settle phase overrun timer
    tonTiming        : TON;    // 计时相正常定时 [TIME] / Timing phase timer
    tonTimingOv      : TON;    // 计时相超时定时 [TIME] / Timing phase overrun timer
    tonRepress       : TON;    // 复压相正常定时 [TIME] / Repressurisation phase timer
    tonRepressOv     : TON;    // 复压相超时定时 [TIME] / Repressurisation phase overrun timer
    tonTotal         : TON;    // 整序总超时定时 [TIME] / Whole-sequence total timeout timer
    rtStart          : R_TRIG; // 启动上升沿检测 [bool] / Start rising edge detector
    rtReset          : R_TRIG; // 复位上升沿检测 [bool] / Reset rising edge detector
    _eState          : E_DL_LyoPrTestState := E_DL_LyoPrTestState.eLyoPrIdle;   // 内部相位（CASE 唯一写入目标）
    _fPressStartMbar : REAL := 0.0;   // 计时相起点压力快照 [mbar] / Base pressure captured at timing start
    _fLeakRaw        : REAL := 0.0;   // 钳制前的原始泄漏率 [mbar*L/s] / Raw leak rate before limiting [mbar*L/s]
    _tElapsed        : TIME := T#0S;  // 计时相实际经过时间 [TIME] / Actual elapsed timing phase duration [TIME]
    _fElapsedS       : REAL := 0.0;   // 计时相实际经过时间折算 [s] / Elapsed timing duration in seconds [s]
    _bFinOk          : BOOL := FALSE; // 实值入参有限性总闸结果 / Finiteness gate aggregate result
    _bVacOk          : BOOL := FALSE; // 起始真空度达成 [bool] / Base vacuum reached flag [bool]
    _bActive         : BOOL := FALSE; // 测试序激活（隔离至复压四相之一）[bool] / Sequence active flag [bool]
    _bPassL          : BOOL := FALSE; // 合格位锁存（跨相保持）[bool] / Pass latch held across phases [bool]
    _bDoneL          : BOOL := FALSE; // 完成位锁存（跨相保持）[bool] / Done latch held across phases [bool]
    _bFault          : BOOL := FALSE; // 故障锁存位 [bool] / Latched fault flag [bool]
    _uInfo           : UDINT := 16#0000_0000;   // 信息码，每拍重算 / Info code, recomputed every cycle
    _uFault          : UDINT := 16#0000_0000;   // 故障码锁存 / Latched fault code
END_VAR
VAR CONSTANT
    DL_EPS         : REAL := 1.0E-9;      // 数值零闸阈值 [-] / Numeric zero gate threshold [-]
    DL_BIG         : REAL := 1.0E12;      // 非有限值闸量级上限 [-] / Finiteness gate magnitude [-]
    DL_VAC_MIN     : REAL := 1.0;         // 起始真空度门槛（压力须低于此值）[mbar] / Base vacuum pressure ceiling [mbar]
    DL_OVER_MARGIN : TIME := T#30S;       // 相超时相对正常定时的裕量 [TIME] / Phase overrun margin [TIME]
    DL_ISO_MAX     : TIME := T#20S;       // 隔离阀动作窗口 [TIME] / Isolation valve travel window [TIME]
    DL_TOTAL_MAX   : TIME := T#2H;        // 整序总超时上限 [TIME] / Whole-sequence total timeout [TIME]
    DL_MS_PER_S    : REAL := 1000.0;      // 毫秒到秒的折算 [ms/s] / Milliseconds per second [ms/s]
    DL_LEAK_HI     : REAL := 100.0;       // 泄漏率物理上限 [mbar*L/s] / Leak rate physical upper bound [mbar*L/s]
END_VAR

(* —— 段 0：单拍量预清零（锁存量 _uFault/_bFault/_bPassL/_bDoneL/_eStatePrev 不入清单，R187①） —— *)
_uInfo := 16#0000_0000;                     // 信息码每拍重算 / Info code recomputed
nErrId := 16#0000_0000;                     // 事件码缺省无事件 / Event code defaults to none

(* —— 段 1：非有限值闸（R19：不拿 NaN 去比较真空度） —— *)
_bFinOk := (fChamberPressMbar > -DL_BIG) AND (fChamberPressMbar < DL_BIG)
           AND (fVolumeL > -DL_BIG) AND (fVolumeL < DL_BIG)
           AND (fLeakMaxMbarLs > -DL_BIG) AND (fLeakMaxMbarLs < DL_BIG);

(* —— 段 2：派生态（真空度达成、序激活、计时换算） —— *)
_bVacOk := _bFinOk AND (fChamberPressMbar <= DL_VAC_MIN);      // 压力低于门槛才算达起始真空
_bActive := (_eState = E_DL_LyoPrTestState.eLyoPrIsolate)
            OR (_eState = E_DL_LyoPrTestState.eLyoPrSettle)
            OR (_eState = E_DL_LyoPrTestState.eLyoPrTiming)
            OR (_eState = E_DL_LyoPrTestState.eLyoPrRepress);
_tElapsed := tonTiming.ET;                                     // 计时相已运行时间（读上拍值，安全）
_fElapsedS := TIME_TO_REAL(_tElapsed) / DL_MS_PER_S;           // 毫秒数折算为秒 [s]（单点赋值，R26）

(* —— 段 3：定时器与边沿无条件周期刷新（R7：调用语句不得置于 IF/CASE 内） —— *)
rtStart(CLK := xStart);                                                                 // 启动上升沿，每拍必调
rtReset(CLK := xReset);                                                                 // 复位上升沿，每拍必调
tonIso(IN := (_eState = E_DL_LyoPrTestState.eLyoPrIsolate), PT := DL_ISO_MAX);          // 隔离相阀动作窗口
tonIsoOv(IN := (_eState = E_DL_LyoPrTestState.eLyoPrIsolate), PT := DL_ISO_MAX + DL_OVER_MARGIN);  // 隔离相超时点
tonSettle(IN := (_eState = E_DL_LyoPrTestState.eLyoPrSettle), PT := tSettleS);          // 稳压相正常定时
tonSettleOv(IN := (_eState = E_DL_LyoPrTestState.eLyoPrSettle),
            PT := tSettleS + DL_OVER_MARGIN);                                           // 稳压相超时点
tonTiming(IN := (_eState = E_DL_LyoPrTestState.eLyoPrTiming), PT := tTestS);            // 计时相正常定时
tonTimingOv(IN := (_eState = E_DL_LyoPrTestState.eLyoPrTiming),
            PT := tTestS + DL_OVER_MARGIN);                                             // 计时相超时点
tonRepress(IN := (_eState = E_DL_LyoPrTestState.eLyoPrRepress), PT := tRepressS);       // 复压相正常定时
tonRepressOv(IN := (_eState = E_DL_LyoPrTestState.eLyoPrRepress),
             PT := tRepressS + DL_OVER_MARGIN);                                         // 复压相超时点
tonTotal(IN := _bActive, PT := DL_TOTAL_MAX);                                           // 整序总超时

(* —— 段 4：全局故障拦截（优先级最高；已锁存则不再改写码值，禁同拍抹除） —— *)
IF xFault AND (NOT _bFault) THEN
    _uFault := 16#0091_0227;                // 故障级：外部故障输入
    _bFault := TRUE;                        // 锁存（3 行内置，R45 配对）
    _eState := E_DL_LyoPrTestState.eLyoPrFault;
END_IF
IF (NOT _bFinOk) AND (NOT _bFault) THEN
    _uFault := 16#0091_0228;                // 故障级：入参非有限
    _bFault := TRUE;                        // 锁存
    _eState := E_DL_LyoPrTestState.eLyoPrFault;
END_IF
IF tonTotal.Q AND _bActive AND (NOT _bFault) THEN
    _uFault := 16#0091_0226;                // 故障级：整序总超时
    _bFault := TRUE;                        // 锁存
    _eState := E_DL_LyoPrTestState.eLyoPrFault;
END_IF

(* —— 段 5：相位机（只做迁移与锁存；出口在段 7 单点映射） —— *)
CASE _eState OF

E_DL_LyoPrTestState.eLyoPrIdle:
    IF NOT xStart THEN
        _bDoneL := FALSE;                   // 撤令即清完成位，为下次测试重新武装
        _bPassL := FALSE;                   // 合格位一并清
    ELSIF NOT _bVacOk THEN
        _uInfo := 16#0091_0221;             // 信息级：未达起始真空度，禁止启动（不置故障位）
    ELSIF rtStart.Q THEN
        _bDoneL := FALSE;                   // 新序开始：清完成位
        _bPassL := FALSE;                   // 新序开始：清合格位
        _eState := E_DL_LyoPrTestState.eLyoPrIsolate;         // 进隔离相
    END_IF

E_DL_LyoPrTestState.eLyoPrIsolate:
    IF NOT xStart THEN
        _uFault := 16#0091_0227;            // 故障级：测试中撤令，按外部中断归因
        _bFault := TRUE;                    // 锁存
        _eState := E_DL_LyoPrTestState.eLyoPrFault;
    ELSIF tonIsoOv.Q THEN
        _uFault := 16#0091_0222;            // 故障级：隔离相超时（隔离阀未关到位）
        _bFault := TRUE;                    // 锁存
        _eState := E_DL_LyoPrTestState.eLyoPrFault;
    ELSIF xIsoValveClosedFb THEN
        _eState := E_DL_LyoPrTestState.eLyoPrSettle;          // 阀关到位：本拍事件优先于超时迁移（R275）
    END_IF

E_DL_LyoPrTestState.eLyoPrSettle:
    IF tonSettleOv.Q THEN
        _uFault := 16#0091_0223;            // 故障级：稳压相超时
        _bFault := TRUE;                    // 锁存
        _eState := E_DL_LyoPrTestState.eLyoPrFault;
    ELSIF tonSettle.Q THEN
        _fPressStartMbar := fChamberPressMbar;                // 计时相起点压力快照（迁移前一次性捕获）
        _eState := E_DL_LyoPrTestState.eLyoPrTiming;          // 进计时相
    END_IF

E_DL_LyoPrTestState.eLyoPrTiming:
    IF tonTimingOv.Q THEN
        _uFault := 16#0091_0224;            // 故障级：计时相超时
        _bFault := TRUE;                    // 锁存
        _eState := E_DL_LyoPrTestState.eLyoPrFault;
    ELSIF tonTiming.Q THEN
        _eState := E_DL_LyoPrTestState.eLyoPrJudge;           // 计时到：进判定相
    END_IF

E_DL_LyoPrTestState.eLyoPrJudge:
    IF (_fElapsedS <= DL_EPS) OR (fVolumeL <= DL_EPS) THEN
        _uFault := 16#0091_0224;            // 故障级：实际计时为零或容积未组态，泄漏率不可算
        _bFault := TRUE;                    // 锁存
        _eState := E_DL_LyoPrTestState.eLyoPrFault;
    ELSE
        _fLeakRaw := (fChamberPressMbar - _fPressStartMbar) * fVolumeL / _fElapsedS;   // 泄漏率 [mbar*L/s]
        IF (_fLeakRaw < 0.0) OR (_fLeakRaw > fLeakMaxMbarLs) THEN
            _uFault := 16#0091_0229;        // 故障级：升压为负（隔离失效）或泄漏率超限
            _bFault := TRUE;                // 锁存
            _eState := E_DL_LyoPrTestState.eLyoPrFault;
        ELSE
            _bPassL := TRUE;                // 合格锁存
            _eState := E_DL_LyoPrTestState.eLyoPrRepress;     // 进复压相
        END_IF
    END_IF

E_DL_LyoPrTestState.eLyoPrRepress:
    IF tonRepressOv.Q THEN
        _uFault := 16#0091_0225;            // 故障级：复压相超时
        _bFault := TRUE;                    // 锁存
        _eState := E_DL_LyoPrTestState.eLyoPrFault;
    ELSIF tonRepress.Q THEN
        _bDoneL := TRUE;                    // 完成位锁存（跨相保持，段 7 单点映射）
        _eState := E_DL_LyoPrTestState.eLyoPrDone;            // 进完成相
    END_IF

E_DL_LyoPrTestState.eLyoPrDone:
    IF xFault THEN
        _uFault := 16#0091_0227;            // 故障级：完成后外部故障（段 4 已拦，此处兜底同码）
        _bFault := TRUE;                    // 锁存
        _eState := E_DL_LyoPrTestState.eLyoPrFault;
    ELSIF NOT xStart THEN
        _bDoneL := FALSE;                   // 撤令：清完成位并回待机
        _eState := E_DL_LyoPrTestState.eLyoPrIdle;
    END_IF

E_DL_LyoPrTestState.eLyoPrFault:
    IF rtReset.Q AND (NOT xFault) AND _bFinOk THEN
        _bFault := FALSE;                   // 解除路径：复位沿 + 外部故障消失 + 入参有限（可达，R188）
        _uFault := 16#0000_0000;            // 清锁存码
        _bDoneL := FALSE;                   // 完成位清
        _bPassL := FALSE;                   // 合格位清，避免故障后误报合格
        _fLeakRaw := 0.0;                   // 泄漏率读数清（故障数据不得留作趋势）
        _eState := E_DL_LyoPrTestState.eLyoPrIdle;            // 回待机，需新上升沿才可再测
    END_IF

ELSE
    _uFault := 16#0091_0230;                // 故障级：非法相位 ID 兜底
    _bFault := TRUE;                        // 锁存
    _eState := E_DL_LyoPrTestState.eLyoPrFault;               // 强制回故障相

END_CASE

(* —— 段 6：后置段（泄漏率读数域兜底：非有限即清零，防污染趋势记录） —— *)
IF NOT (_fLeakRaw > -DL_BIG AND _fLeakRaw < DL_BIG) THEN
    _fLeakRaw := 0.0;                       // 内部状态自检：非有限即清零
END_IF

(* —— 段 7：出口单点映射（名实同源；阀门由状态导出，故障侧一律关阀） —— *)
xIsoValveCmd := ((_eState = E_DL_LyoPrTestState.eLyoPrIsolate)
                 OR (_eState = E_DL_LyoPrTestState.eLyoPrSettle)
                 OR (_eState = E_DL_LyoPrTestState.eLyoPrTiming)
                 OR (_eState = E_DL_LyoPrTestState.eLyoPrJudge)
                 OR (_eState = E_DL_LyoPrTestState.eLyoPrRepress)) AND (NOT _bFault);   // 隔离阀：五相关闭
xVentCmd := (_eState = E_DL_LyoPrTestState.eLyoPrRepress) AND (NOT _bFault);             // 通气阀：仅复压相开
fLeakRateMbarLs := LIMIT(0.0, _fLeakRaw, DL_LEAK_HI);                                    // 泄漏率钳 0..物理上限
xTestPass := _bPassL AND (NOT _bFault);                                                  // 合格位出口
xDone := _bDoneL AND (NOT _bFault);                                                      // 完成位出口
xBusy := _bActive AND (NOT _bFault);                                                     // 进行中出口
eState := _eState;                                                                       // 状态出口单点映射
IF _bFault THEN
    nErrId := _uFault;                      // 故障锁存码回放（不在故障相按当下输入重推断）
ELSE
    nErrId := _uInfo;                       // 信息码
END_IF

END_FUNCTION_BLOCK
